ORGANIZATION_BLOCK "PullOrPlugOfModules"   // OB83, LAD, PullOrPlugOfModules
{ S7_Optimized_Access := 'TRUE' }
VERSION : 0.1
// stored: IsIECCheckEnabled false, SetENOAutomatically false
   VAR_INPUT
      LADDR : HW_IO;   // Hardware identifier
      Event_Class : Byte;   // 16#38/39: module inserted, removed
      Fault_ID : Byte;   // Fault identifier
   END_VAR
BEGIN
END_ORGANIZATION_BLOCK

ORGANIZATION_BLOCK "RackOrStationFailure"   // OB86, LAD, RackOrStationFailure
{ S7_Optimized_Access := 'TRUE' }
VERSION : 0.1
// stored: IsIECCheckEnabled false, SetENOAutomatically false
   VAR_INPUT
      LADDR : HW_DEVICE;   // Hardware identifier
      Event_Class : Byte;   // Event class
      Fault_ID : Byte;   // Fault identifier
   END_VAR
BEGIN
END_ORGANIZATION_BLOCK

FUNCTION "ByteArrayToString" : String   // FC15, SCL
{ S7_Optimized_Access := 'TRUE' }
VERSION : 0.1
// stored: AutoNumber true, IsIECCheckEnabled false, SetENOAutomatically false, UDAEnableTagReadback false
   VAR_INPUT
      Lenght : Int;
      ByteArray : Array[0..1024] of Byte;
   END_VAR
   VAR_OUTPUT
      ByteArrayToString_1 : String;
      ByteArrayToString_2 : String;
      ByteArrayToString_3 : String;
      ByteArrayToString_4 : String;
      ByteArrayToString_5 : String;
   END_VAR
   VAR_TEMP
      tempStr_1 : String;
      tempStr_2 : String;
      tempStr_3 : String;
      tempStr_4 : String;
      tempStr_5 : String;
      tempStr_6 : String;
      foundPos : Int;
      i : Int;
   END_VAR
BEGIN
   //STRING 1
   #tempStr_1 := '';
   FOR #i := 0 TO MIN(IN1 := #Lenght - 1, IN2 := 254) DO
       IF #ByteArray[#i] <> 0 THEN
           #tempStr_1 := CONCAT(IN1 := #tempStr_1, IN2 := CHAR_TO_STRING(BYTE_TO_CHAR(#ByteArray[#i])));
       END_IF;
   END_FOR;

   //STRING 2
   #tempStr_2 := '';
   FOR #i := 100 TO MIN(IN1 := #Lenght - 1, IN2 := 354) DO
       IF #ByteArray[#i] <> 0 THEN
           #tempStr_2 := CONCAT(IN1 := #tempStr_2, IN2 := CHAR_TO_STRING(BYTE_TO_CHAR(#ByteArray[#i])));
       END_IF;
   END_FOR;

   //STRING 3
   #tempStr_3 := '';
   FOR #i := 200 TO MIN(IN1 := #Lenght - 1, IN2 := 454) DO
       IF #ByteArray[#i] <> 0 THEN
           #tempStr_3 := CONCAT(IN1 := #tempStr_3, IN2 := CHAR_TO_STRING(BYTE_TO_CHAR(#ByteArray[#i])));
       END_IF;
   END_FOR;

   //STRING 4
   #tempStr_4 := '';
   FOR #i := 300 TO MIN(IN1 := #Lenght - 1, IN2 := 554) DO
       IF #ByteArray[#i] <> 0 THEN
           #tempStr_4 := CONCAT(IN1 := #tempStr_4, IN2 := CHAR_TO_STRING(BYTE_TO_CHAR(#ByteArray[#i])));
       END_IF;
   END_FOR;

   // //STRING 5
   #tempStr_5 := '';
   FOR #i := 400 TO MIN(IN1 := #Lenght - 1, IN2 := 654) DO
       IF #ByteArray[#i] <> 0 THEN
           #tempStr_5 := CONCAT(IN1 := #tempStr_5, IN2 := CHAR_TO_STRING(BYTE_TO_CHAR(#ByteArray[#i])));
       END_IF;
   END_FOR;

   // //STRING 6
   #tempStr_6 := '';
   FOR #i := 500 TO MIN(IN1 := #Lenght - 1, IN2 := 763) DO
       IF #ByteArray[#i] <> 0 THEN
           #tempStr_6 := CONCAT(IN1 := #tempStr_6, IN2 := CHAR_TO_STRING(BYTE_TO_CHAR(#ByteArray[#i])));
       END_IF;
   END_FOR;

   // Remove '$R$L'
   // string 1
   #foundPos := FIND(IN1 := #tempStr_1, IN2 := '$R$L');
   WHILE #foundPos > 0 DO
       #tempStr_1 := REPLACE(IN1 := #tempStr_1, IN2 := '', P := #foundPos, L := 2);
       #foundPos := FIND(IN1 := #tempStr_1, IN2 := '$R$L');
   END_WHILE;

   // string 2
   #foundPos := FIND(IN1 := #tempStr_2, IN2 := '$R$L');
   WHILE #foundPos > 0 DO
       #tempStr_2 := REPLACE(IN1 := #tempStr_2, IN2 := '', P := #foundPos, L := 2);
       #foundPos := FIND(IN1 := #tempStr_2, IN2 := '$R$L');
   END_WHILE;

   // string 3
   #foundPos := FIND(IN1 := #tempStr_3, IN2 := '$R$L');
   WHILE #foundPos > 0 DO
       #tempStr_3 := REPLACE(IN1 := #tempStr_3, IN2 := '', P := #foundPos, L := 2);
       #foundPos := FIND(IN1 := #tempStr_3, IN2 := '$R$L');
   END_WHILE;

   // string 4
   #foundPos := FIND(IN1 := #tempStr_4, IN2 := '$R$L');
   WHILE #foundPos > 0 DO
       #tempStr_4 := REPLACE(IN1 := #tempStr_4, IN2 := '', P := #foundPos, L := 2);
       #foundPos := FIND(IN1 := #tempStr_4, IN2 := '$R$L');
   END_WHILE;

   // string 5
   #foundPos := FIND(IN1 := #tempStr_5, IN2 := '$R$L');
   WHILE #foundPos > 0 DO
       #tempStr_5 := REPLACE(IN1 := #tempStr_5, IN2 := '', P := #foundPos, L := 2);
       #foundPos := FIND(IN1 := #tempStr_5, IN2 := '$R$L');
   END_WHILE;

   // string 6
   #foundPos := FIND(IN1 := #tempStr_6, IN2 := '$R$L');
   WHILE #foundPos > 0 DO
       #tempStr_6 := REPLACE(IN1 := #tempStr_6, IN2 := '', P := #foundPos, L := 2);
       #foundPos := FIND(IN1 := #tempStr_6, IN2 := '$R$L');
   END_WHILE;

   #ByteArrayToString := #tempStr_1;
   #ByteArrayToString_1 := #tempStr_2;
   #ByteArrayToString_2 := #tempStr_3;
   #ByteArrayToString_3 := #tempStr_4;
   #ByteArrayToString_4 := #tempStr_5;
   #ByteArrayToString_5 := #tempStr_6;
END_FUNCTION

FUNCTION "ByteArrayToString_1" : String   // FC23, SCL
{ S7_Optimized_Access := 'TRUE' }
VERSION : 0.1
// stored: AutoNumber true, IsIECCheckEnabled false, SetENOAutomatically false, UDAEnableTagReadback false
   VAR_INPUT
      Lenght : Int;
      ByteArray : Array[1..200] of Byte;
   END_VAR
   VAR_TEMP
      tempStr_1 : String;
      foundPos : Int;
      i : Int;
   END_VAR
BEGIN
   #tempStr_1 := '';
   FOR #i := 1 TO MIN(IN1 := #Lenght - 1, IN2 := 200) DO
       IF #ByteArray[#i] <> 0 THEN
           #tempStr_1 := CONCAT(IN1 := #tempStr_1, IN2 := CHAR_TO_STRING(BYTE_TO_CHAR(#ByteArray[#i])));
       END_IF;
   END_FOR;

   // Remove '$02'
   // string 1
   #foundPos := FIND(IN1 := #tempStr_1, IN2 := '$02');
   WHILE #foundPos > 0 DO
       #tempStr_1 := REPLACE(IN1 := #tempStr_1, IN2 := '', P := #foundPos, L := 1);
       #foundPos := FIND(IN1 := #tempStr_1, IN2 := '$02');
   END_WHILE;

   #ByteArrayToString_1 := #tempStr_1;
END_FUNCTION

FUNCTION "CharsArrayToString" : String   // FC27, SCL
{ S7_Optimized_Access := 'TRUE' }
VERSION : 0.1
// stored: AutoNumber true, IsIECCheckEnabled false, SetENOAutomatically false, UDAEnableTagReadback false
   VAR_INPUT
      Lenght : Int;
      CharsArray : Array[1..16] of Char;
   END_VAR
   VAR_TEMP
      tempStr_1 : String;
      foundPos : Int;
      i : Int;
   END_VAR
BEGIN
   #tempStr_1 := '';
   FOR #i := 1 TO MIN(IN1 := #Lenght - 1, IN2 := 16) DO
       IF #CharsArray[#i] <> '$00' THEN
           #tempStr_1 := CONCAT(IN1 := #tempStr_1, IN2 := CHAR_TO_STRING(#CharsArray[#i]));
       END_IF;
   END_FOR;

   // Remove '$00'
   // string 1
   #foundPos := FIND(IN1 := #tempStr_1, IN2 := '$00');
   WHILE #foundPos > 0 DO
       #tempStr_1 := REPLACE(IN1 := #tempStr_1, IN2 := '', P := #foundPos, L := 1);
       #foundPos := FIND(IN1 := #tempStr_1, IN2 := '$00');
   END_WHILE;

   #CharsArrayToString := #tempStr_1;
END_FUNCTION

FUNCTION "FindBoolField" : Bool   // FC17, SCL
{ S7_Optimized_Access := 'TRUE' }
VERSION : 0.1
// stored: AutoNumber true, IsIECCheckEnabled false, SetENOAutomatically false, UDAEnableTagReadback false
   VAR_INPUT
      FieldName : String;
      JsonStr : String;
   END_VAR
   VAR_TEMP
      searchStr : String;
      foundPos : Int;
      valueStr : String;
      afterField : String;
      bResult : Bool;
   END_VAR
BEGIN
   // Build search string
   #searchStr := CONCAT(IN1 := '"', IN2 := #FieldName);
   #searchStr := CONCAT(IN1 := #searchStr, IN2 := '" :');

   // Serach for JSON field
   #foundPos := FIND(IN1 := #JsonStr, IN2 := #searchStr);

   IF #foundPos > 0 THEN
       // Take to 20 characters after the field
       #afterField := MID(IN := #JsonStr, P := #foundPos + LEN(#searchStr), L := 20);

       // Normalize to remove whitespace if necessary
       // (or compare directly)
       IF FIND(IN1 := #afterField, IN2 := 'true') > 0 THEN
           #bResult := TRUE;
       ELSIF FIND(IN1 := #afterField, IN2 := 'false') > 0 THEN
           #bResult := FALSE;
       ELSE
           #bResult := FALSE; // default if value not found
       END_IF;
   ELSE
       #bResult := FALSE;
   END_IF;

   #FindBoolField := #bResult;
END_FUNCTION

FUNCTION "FindDINTFieldFragmented" : DInt   // FC20, SCL
{ S7_Optimized_Access := 'TRUE' }
VERSION : 0.1
// stored: AutoNumber true, IsIECCheckEnabled false, SetENOAutomatically false, UDAEnableTagReadback false
   VAR_INPUT
      FieldName : String;
      Str1 : String;
      Str2 : String;
   END_VAR
   VAR_TEMP
      searchStr : String;
      iStart : Int;
      iEnd : Int;
      tempVal : String;
      fieldFound : Bool;
      loopIdx : Int;
   END_VAR
BEGIN
   // Build search string
   #searchStr := CONCAT(IN1 := '"', IN2 := #FieldName);
   #searchStr := CONCAT(IN1 := #searchStr, IN2 := '" :');

   // Serach for JSON field
   #iStart := FIND(IN1 := #Str1, IN2 := #searchStr);

   IF #iStart > 0 THEN
       // Found full field in String_1
       #iEnd := FIND(IN1 := MID(IN := #Str1, P := #iStart + LEN(#searchStr), L := 20), IN2 := ',');
       IF #iEnd = 0 THEN
           #iEnd := FIND(IN1 := MID(IN := #Str1, P := #iStart + LEN(#searchStr), L := 20), IN2 := '}');
       END_IF;
       IF #iEnd > 0 THEN
           #tempVal := MID(IN := #Str1, P := #iStart + LEN(#searchStr), L := #iEnd - 1);
           #fieldFound := TRUE;
       END_IF;
   END_IF;

   // Search for full field in Str2
   IF NOT #fieldFound THEN
       #iStart := FIND(IN1 := #Str2, IN2 := #searchStr);
       IF #iStart > 0 THEN
           #iEnd := FIND(IN1 := MID(IN := #Str2, P := #iStart + LEN(#searchStr), L := 20), IN2 := ',');
           IF #iEnd = 0 THEN
               #iEnd := FIND(IN1 := MID(IN := #Str2, P := #iStart + LEN(#searchStr), L := 20), IN2 := '}');
           END_IF;
           IF #iEnd > 0 THEN
               #tempVal := MID(IN := #Str2, P := #iStart + LEN(#searchStr), L := #iEnd - 1);
               #fieldFound := TRUE;
           END_IF;
       END_IF;
   END_IF;

   // Search for fragmented field: end of name in Str1 and beginning in Str2
   IF NOT #fieldFound THEN
       // Examines last 10 characters of String_1
       FOR #loopIdx := LEN(#Str1) - 15 TO LEN(#Str1) DO
           IF MID(IN := #Str1, P := #loopIdx, L := 1) = '"' THEN
               #tempVal := MID(IN := #Str1, P := #loopIdx, L := LEN(#Str1) - #loopIdx + 1);
               #tempVal := CONCAT(IN1 := #tempVal, IN2 := #Str2); // concatenates piece from beginning of String_2
               #iStart := FIND(IN1 := #tempVal, IN2 := #searchStr);
               IF #iStart > 0 THEN
                   #iEnd := FIND(IN1 := MID(IN := #tempVal, P := #iStart + LEN(#searchStr), L := 20), IN2 := ',');
                   IF #iEnd = 0 THEN
                       #iEnd := FIND(IN1 := MID(IN := #tempVal, P := #iStart + LEN(#searchStr), L := 20), IN2 := '}');
                   END_IF;
                   IF #iEnd > 0 THEN
                       #tempVal := MID(IN := #tempVal, P := #iStart + LEN(#searchStr), L := #iEnd - 1);
                       #fieldFound := TRUE;
                   END_IF;
               END_IF;
               EXIT; // found, you can leave
           END_IF;
       END_FOR;
   END_IF;

   // Return value
   IF #fieldFound THEN
       #FindDINTFieldFragmented := STRING_TO_DINT(#tempVal);
   ELSE
       #FindDINTFieldFragmented := -9999; // default value if not found
   END_IF;
END_FUNCTION

FUNCTION "FindINTFieldFragmented" : Int   // FC22, SCL
{ S7_Optimized_Access := 'TRUE' }
VERSION : 0.1
// stored: AutoNumber true, IsIECCheckEnabled false, SetENOAutomatically false, UDAEnableTagReadback false
   VAR_INPUT
      FieldName : String;
      Str1 : String;
      Str2 : String;
   END_VAR
   VAR_TEMP
      searchStr : String;
      iStart : Int;
      iEnd : Int;
      tempVal : String;
      fieldFound : Bool;
      loopIdx : Int;
   END_VAR
BEGIN
   // Build search string
   #searchStr := CONCAT(IN1 := '"', IN2 := #FieldName);
   #searchStr := CONCAT(IN1 := #searchStr, IN2 := '" :');

   // Serach for JSON field
   #iStart := FIND(IN1 := #Str1, IN2 := #searchStr);

   IF #iStart > 0 THEN
       // Found full field in String_1
       #iEnd := FIND(IN1 := MID(IN := #Str1, P := #iStart + LEN(#searchStr), L := 20), IN2 := ',');
       IF #iEnd = 0 THEN
           #iEnd := FIND(IN1 := MID(IN := #Str1, P := #iStart + LEN(#searchStr), L := 20), IN2 := '}');
       END_IF;
       IF #iEnd > 0 THEN
           #tempVal := MID(IN := #Str1, P := #iStart + LEN(#searchStr), L := #iEnd - 1);
           #fieldFound := TRUE;
       END_IF;
   END_IF;

   // Search for full field in Str2
   IF NOT #fieldFound THEN
       #iStart := FIND(IN1 := #Str2, IN2 := #searchStr);
       IF #iStart > 0 THEN
           #iEnd := FIND(IN1 := MID(IN := #Str2, P := #iStart + LEN(#searchStr), L := 20), IN2 := ',');
           IF #iEnd = 0 THEN
               #iEnd := FIND(IN1 := MID(IN := #Str2, P := #iStart + LEN(#searchStr), L := 20), IN2 := '}');
           END_IF;
           IF #iEnd > 0 THEN
               #tempVal := MID(IN := #Str2, P := #iStart + LEN(#searchStr), L := #iEnd - 1);
               #fieldFound := TRUE;
           END_IF;
       END_IF;
   END_IF;

   // Search for fragmented field: end of name in Str1 and beginning in Str2
   IF NOT #fieldFound THEN
       // Examines last 10 characters of String_1
       FOR #loopIdx := LEN(#Str1) - 15 TO LEN(#Str1) DO
           IF MID(IN := #Str1, P := #loopIdx, L := 1) = '"' THEN
               #tempVal := MID(IN := #Str1, P := #loopIdx, L := LEN(#Str1) - #loopIdx + 1);
               #tempVal := CONCAT(IN1 := #tempVal, IN2 := #Str2); // concatenates piece from beginning of String_2
               #iStart := FIND(IN1 := #tempVal, IN2 := #searchStr);
               IF #iStart > 0 THEN
                   #iEnd := FIND(IN1 := MID(IN := #tempVal, P := #iStart + LEN(#searchStr), L := 20), IN2 := ',');
                   IF #iEnd = 0 THEN
                       #iEnd := FIND(IN1 := MID(IN := #tempVal, P := #iStart + LEN(#searchStr), L := 20), IN2 := '}');
                   END_IF;
                   IF #iEnd > 0 THEN
                       #tempVal := MID(IN := #tempVal, P := #iStart + LEN(#searchStr), L := #iEnd - 1);
                       #fieldFound := TRUE;
                   END_IF;
               END_IF;
               EXIT; // found, you can leave
           END_IF;
       END_FOR;
   END_IF;

   // Return value
   IF #fieldFound THEN
       #FindINTFieldFragmented := STRING_TO_INT(#tempVal);
   ELSE
       #FindINTFieldFragmented := -9999; // default value if not found
   END_IF;
END_FUNCTION

FUNCTION "FindIntField" : Int   // FC18, SCL
{ S7_Optimized_Access := 'TRUE' }
VERSION : 0.1
// stored: AutoNumber true, IsIECCheckEnabled false, SetENOAutomatically false, UDAEnableTagReadback false
   VAR_INPUT
      FieldName : String;
      JsonStr : String;
   END_VAR
   VAR_TEMP
      searchStr : String;
      foundPos : Int;
      valueStr : String;
      delimPos : Int;
   END_VAR
BEGIN
   // Set up the search pattern, e.g. '"id":'
   #searchStr := CONCAT(IN1 := '"', IN2 := #FieldName);
   #searchStr := CONCAT(IN1 := #searchStr, IN2 := '" :');

   // Search the field
   #foundPos := FIND(IN1 := #JsonStr, IN2 := #searchStr);

   IF #foundPos > 0 THEN
       // Try to find a comma after the value
       #delimPos := FIND(
                         IN1 := MID(IN := #JsonStr, P := #foundPos + LEN(#searchStr), L := 10),
                         IN2 := ','
       );

       // If there is no comma, try to find the closing brace '}'
       IF #delimPos = 0 THEN
           #delimPos := FIND(
                             IN1 := MID(IN := #JsonStr, P := #foundPos + LEN(#searchStr), L := 10),
                             IN2 := '}'
           );
       END_IF;

       // If you find the end of value, extract the value
       IF #delimPos > 0 THEN
           #valueStr := MID(
                            IN := #JsonStr,
                            P := #foundPos + LEN(#searchStr),
                            L := #delimPos - 1
           );
           #FindIntField := STRING_TO_INT(#valueStr);
           RETURN;
       END_IF;
   END_IF;

   // Default return if not found or error
   #FindIntField := -9999;
END_FUNCTION

FUNCTION "FindSTRINGFieldFragmented" : String   // FC21, SCL
{ S7_Optimized_Access := 'TRUE' }
VERSION : 0.1
// stored: AutoNumber true, IsIECCheckEnabled false, SetENOAutomatically false, UDAEnableTagReadback false
   VAR_INPUT
      FieldName : String;
      Str1 : String;
      Str2 : String;
   END_VAR
   VAR_TEMP
      searchStr : String;
      iStart : Int;
      iEnd : Int;
      tempVal : String;
      fieldFound : Bool;
      loopIdx : Int;
   END_VAR
BEGIN
   // Build search string
   #searchStr := CONCAT(IN1 := '"', IN2 := #FieldName);
   #searchStr := CONCAT(IN1 := #searchStr, IN2 := '" :');

   // Serach for JSON field
   #iStart := FIND(IN1 := #Str1, IN2 := #searchStr);

   IF #iStart > 0 THEN
       // Found full field in String_1
       #iEnd := FIND(IN1 := MID(IN := #Str1, P := #iStart + LEN(#searchStr), L := 20), IN2 := ',');
       IF #iEnd = 0 THEN
           #iEnd := FIND(IN1 := MID(IN := #Str1, P := #iStart + LEN(#searchStr), L := 20), IN2 := '}');
       END_IF;
       IF #iEnd > 0 THEN
           #tempVal := MID(IN := #Str1, P := #iStart + LEN(#searchStr), L := #iEnd - 1);
           #fieldFound := TRUE;
       END_IF;
   END_IF;

   // Search for full field in Str2
   IF NOT #fieldFound THEN
       #iStart := FIND(IN1 := #Str2, IN2 := #searchStr);
       IF #iStart > 0 THEN
           #iEnd := FIND(IN1 := MID(IN := #Str2, P := #iStart + LEN(#searchStr), L := 20), IN2 := ',');
           IF #iEnd = 0 THEN
               #iEnd := FIND(IN1 := MID(IN := #Str2, P := #iStart + LEN(#searchStr), L := 20), IN2 := '}');
           END_IF;
           IF #iEnd > 0 THEN
               #tempVal := MID(IN := #Str2, P := #iStart + LEN(#searchStr), L := #iEnd - 1);
               #fieldFound := TRUE;
           END_IF;
       END_IF;
   END_IF;

   // Search for fragmented field: end of name in Str1 and beginning in Str2
   IF NOT #fieldFound THEN
       // Examines last 10 characters of String_1
       FOR #loopIdx := LEN(#Str1) - 15 TO LEN(#Str1) DO
           IF MID(IN := #Str1, P := #loopIdx, L := 1) = '"' THEN
               #tempVal := MID(IN := #Str1, P := #loopIdx, L := LEN(#Str1) - #loopIdx + 1);
               #tempVal := CONCAT(IN1 := #tempVal, IN2 := #Str2); // concatenates piece from beginning of String_2
               #iStart := FIND(IN1 := #tempVal, IN2 := #searchStr);
               IF #iStart > 0 THEN
                   #iEnd := FIND(IN1 := MID(IN := #tempVal, P := #iStart + LEN(#searchStr), L := 20), IN2 := ',');
                   IF #iEnd = 0 THEN
                       #iEnd := FIND(IN1 := MID(IN := #tempVal, P := #iStart + LEN(#searchStr), L := 20), IN2 := '}');
                   END_IF;
                   IF #iEnd > 0 THEN
                       #tempVal := MID(IN := #tempVal, P := #iStart + LEN(#searchStr), L := #iEnd - 1);
                       #fieldFound := TRUE;
                   END_IF;
               END_IF;
               EXIT; // found, you can leave
           END_IF;
       END_FOR;
   END_IF;

   // Return value
   IF #fieldFound THEN
       #FindSTRINGFieldFragmented := #tempVal;
   ELSE
       #FindSTRINGFieldFragmented := 'NOT FOUND'; // default value if not found
   END_IF;
END_FUNCTION

FUNCTION "FindStringField" : String   // FC19, SCL
{ S7_Optimized_Access := 'TRUE' }
VERSION : 0.1
// stored: AutoNumber true, IsIECCheckEnabled false, SetENOAutomatically false, UDAEnableTagReadback false
   VAR_INPUT
      FieldName : String;
      JsonStr : String;
   END_VAR
   VAR_TEMP
      searchStr : String;
      foundPos : Int;
      resultStr : String;
      quotePos1 : Int;
      quotePos2 : Int;
   END_VAR
BEGIN
   // Sets search pattern → ex: '"loadstate":'
   #searchStr := CONCAT(IN1 := '"', IN2 := #FieldName);
   #searchStr := CONCAT(IN1 := #searchStr, IN2 := '" :');

   // Search in JSON
   #foundPos := FIND(IN1 := #JsonStr, IN2 := #searchStr);

   IF #foundPos > 0 THEN
       // Finds first quote after field
       #quotePos1 := FIND(IN1 := MID(IN := #JsonStr, P := #foundPos + LEN(#searchStr), L := 20), IN2 := '"');

       IF #quotePos1 > 0 THEN
           // Finds second quote after the first
           #quotePos2 := FIND(
                              IN1 := MID(IN := #JsonStr, P := #foundPos + LEN(IN := #searchStr) + #quotePos1, L := 10),
                              IN2 := '"'
           );

           IF #quotePos2 > 0 THEN
               #resultStr := MID(
                                 IN := #JsonStr,
                                 P := #foundPos + LEN(#searchStr) + #quotePos1,
                                 L := #quotePos2 - 1
               );
               #FindStringField := #resultStr;
               RETURN;
           END_IF;
       END_IF;
   END_IF;

   // If not found, returns empty string
   #FindStringField := '';
END_FUNCTION

FUNCTION "ID_Decode_F" : Void   // FC3, SCL
{ S7_Optimized_Access := 'TRUE' }
VERSION : 0.1
// stored: AutoNumber true, IsIECCheckEnabled false, SetENOAutomatically false, UDAEnableTagReadback false
   VAR_INPUT
      ID : DInt;
   END_VAR
   VAR_IN_OUT
      ID_Decoded : "ID_Decoded";
   END_VAR
   VAR_TEMP
      Temp : UInt;
   END_VAR
BEGIN

   // Extract XX (first two digits)
   #ID_Decoded.Device_Type := #ID / 10000;        // 123456 / 10000 = 12

   // Extract YY (middle two digits)
   #ID_Decoded.Level := (#ID MOD 10000) / 100; // 123456 % 10000 = 3456 → 3456 / 100 = 34

   // Extract ZZ (last two digits)
   #ID_Decoded.VTD := #ID MOD 100;       // 123456 % 100 = 56
END_FUNCTION

FUNCTION "IsIPAddress" : Bool   // FC4, SCL
TITLE = IsIPAddress
{ S7_Optimized_Access := 'TRUE' }
VERSION : 0.1
// Evaluates whether a given String contains a valid IP address
// stored: AutoNumber true, IsIECCheckEnabled true, SetENOAutomatically true, UDAEnableTagReadback false
   VAR_INPUT
      address : String;   // Address to be evaluated
   END_VAR
   VAR_OUTPUT
      ipAddress : IP_V4;   // Parsed IP address if passed address is IP address
   END_VAR
   VAR_TEMP
      tempAddress : String;   // Passed address
      tempOctet : String;   // Current octet
      tempIndex : DInt;   // Index for loop
      tempPos : Int;   // Position of found separator
      tempNum : Int;   // Converted octet
      tempIp : IP_V4;   // Parsed IP address
   END_VAR
   VAR CONSTANT
      MAX_VALUE : USInt := 255;   // Max. valid value of octet
      NUM_OCTETS : DInt := 4;   // Number of octets
      CHAR_ZERO : Char := '0';   // ASCII character '0'
   END_VAR
   // Ret_Val : Return value
BEGIN
   REGION BLOCK INFO HEADER
     //===============================================================================
     // SIEMENS / (c)Copyright 2024
     //-------------------------------------------------------------------------------
     // Title:        IsIPAddress
     // Function:     Evaluates whether a given String contains a valid IP address
     // Library:      --
     // Author:       Siemens Industry Online Support
     // Tested with:  CPU 1515-2 PN V3.1
     // Engineering:  TIA Portal V17
     // Restrictions: --
     // Requirements: S7-1200 with firmware V4.4 or higher
     //               S7-1500 with firmware V2.0 or higher
     //-------------------------------------------------------------------------------
     // Change log table:
     // Version  | Date       | Expert in charge       | Changes applied
     //-------------------------------------------------------------------------------
     // 01.00.00 | 2024-02-12 | Online Support         | First released version
     //===============================================================================
   END_REGION

   #tempAddress := #address;
   #IsIPAddress := FALSE; // Will be overwritten if IP address is detected
   #ipAddress := #tempIp; // Zero output parameter

   FOR #tempIndex := 1 TO #NUM_OCTETS DO
     #tempPos := FIND(IN1 := #tempAddress, IN2 := '.'); // Find separator

     IF (#tempPos > 0 OR #tempIndex = #NUM_OCTETS) // Separator found with exception of last octet
       AND NOT (#tempPos > 0 AND #tempIndex = #NUM_OCTETS) // No separator found in last octet
       AND #tempPos <= 4 // 3  characters or less
     THEN
       IF #tempIndex < #NUM_OCTETS THEN // First three octets
         #tempOctet := LEFT(IN := #tempAddress, L := #tempPos - 1);
       ELSE// Last octet
         #tempOctet := #tempAddress;
       END_IF;

       STRG_VAL(IN := #tempOctet,
                FORMAT := 0,
                P := 1,
                OUT => #tempNum);

       IF #tempNum >= 0 AND #tempNum <= #MAX_VALUE // Within 0 and 255
         AND NOT (#tempNum = 0 AND #tempIndex = 1) // Not 0 in first octet
         AND NOT (#tempNum = 0 AND #tempOctet[1] <> #CHAR_ZERO) // Not 0 because of invalid character
       THEN
         #tempIp.ADDR[#tempIndex] := INT_TO_BYTE(#tempNum);
         #tempAddress := RIGHT(IN := #tempAddress, L := LEN(#tempAddress) - #tempPos); // Remove evaluated octet
       ELSE // Address is not IP address
         EXIT;
       END_IF;
     ELSE // Address is not IP address
       EXIT;
     END_IF;

     IF #tempIndex = #NUM_OCTETS THEN // End of loop reached, address is IP address
       #ipAddress := #tempIp;
       #IsIPAddress := true;
     END_IF;
   END_FOR;
END_FUNCTION

FUNCTION "LMQTT_ConvertToUtf8" : Void   // FC6, SCL
TITLE = LMQTT_ConvertToUtf8
{ S7_Optimized_Access := 'TRUE' }
AUTHOR : SIEMENS
FAMILY : LMQTT
VERSION : 1.0
// Function to convert a WCHAR to a UTF-8 conformant byte sequence
// stored: AutoNumber true, IsIECCheckEnabled true, SetENOAutomatically false, UDAEnableTagReadback false
   VAR_INPUT
      character : WChar;   // Character that shall be converted to UTF-8
   END_VAR
   VAR_OUTPUT
      convertedUtf8 : DWord;   // UTF-8 conformant byte sequence. B0 stores first Byte, B1 second and B2 third Byte. B3 is not used
      bytesUsed : USInt;   // Amount of Bytes converted. Ranges from 1 to 3.
      error : Bool;   // TRUE: An error occurred during the execution of the FC
      status : Word;   // 16#0000 - 16#7FFF: Status of the FC, 16#8000 - 16#FFFF: Error identification
   END_VAR
   VAR_TEMP
      tempStatus : Word;   // temp value for output 'status'
      tempConvertedUtf8 : DWord;   // temp value for output 'convertedUtf8'
      tempBytesUsed : USInt;   // temp value for output 'bytesUsed'
      tempCharacter : WChar;   // temp value for input 'character'
   END_VAR
   VAR CONSTANT
      STATUS_NO_ERROR : Word := 16#0000;   // no error status
      STATUS_EXECUTION_FINISHED : Word := 16#0000;   // Execution finished without errors
      ERR_UNDEFINED : Word := 16#8000;   // Error due to an undefined case
      USINT_NULL : USInt := 0;   // Init value with 0
      DWORD_NULL : DWord := 16#0000_0000;   // Init value with 0
      EMPTY_WCHAR : WChar := WCHAR#' ';   // Empty WChar for comparison
      BELOW_7F : Word := 16#007F;   // Upper limit for character if only one Byte used
      BELOW_7FF : Word := 16#07FF;   // Upper limit for character if two Byte used
      BELOW_MAX_FFFF : Word := 16#FFFF;   // Upper limit for character if three Byte used
      BYTE_3F : Byte := 16#3F;   // Conversion Value
      BYTE_80 : Byte := 16#80;   // Conversion Value
      BYTE_C0 : Byte := 16#C0;   // Conversion Value
      BYTE_E0 : Byte := 16#E0;   // Conversion Value
      USINT_ONE : USInt := 1;   // Const Value to assign amount of bytes used
      USINT_TWO : USInt := 2;   // Const Value to assign amount of bytes used
      USINT_THREE : USInt := 3;   // Const Value to assign amount of bytes used
   END_VAR
   // Ret_Val : No return for this FC - see error and status output
BEGIN
   REGION BLOCK INFO HEADER
       //=============================================================================
       // SIEMENS AG
       // (c)Copyright 2020
       //-----------------------------------------------------------------------------
       // Library:       LMQTT
       // Tested with:   CPU 1516-3 PN/DP V2.8
       // Engineering:   TIA Portal V16
       // Restrictions:  --
       // Requirements:  --
       // Functionality: Converts a single WChar Character to a valid UTF-8 encoded byte sequence and saves this to a DWord.
       //                The amount of bytes saved is stored in bytesUsed Output.
       //-----------------------------------------------------------------------------
       // Change log table:
       // Version    Date         Expert in charge         Changes applied
       // 03.00.00   01.10.2020   Siemens Online Support   First released version
       //=============================================================================
   END_REGION

   REGION INITIALISATION  
       // Initialize functionality: reset of variables, diagnostics, etc.
       #tempConvertedUtf8 := #DWORD_NULL;
       #tempBytesUsed := #USINT_NULL;
       #tempStatus := #STATUS_NO_ERROR;
       //assign temp value from input:
        #tempCharacter := #character;

   END_REGION

   REGION PROGRAM LOGIC
       // Use this region for application specific code
       IF #tempCharacter = #EMPTY_WCHAR THEN
           //will be only 1 byte occupied
           #tempConvertedUtf8 := WCHAR_TO_DWORD(#tempCharacter);
           #tempBytesUsed := #USINT_ONE;
       ELSIF (WCHAR_TO_WORD(#tempCharacter) <= (#BELOW_7F)) THEN
           //will be only 1 byte occupied
           #tempConvertedUtf8 := WCHAR_TO_DWORD(#tempCharacter);
           #tempBytesUsed := #USINT_ONE;
       ELSIF (WCHAR_TO_WORD(#tempCharacter) <= (#BELOW_7FF)) THEN
           //will be 2 byte occupied
           #tempConvertedUtf8.%B1 := (WCHAR_TO_BYTE(#tempCharacter) AND #BYTE_3F) OR #BYTE_80;
           #tempConvertedUtf8.%B0 := WORD_TO_BYTE(SHR(IN := WCHAR_TO_WORD(#tempCharacter), N := 6)) OR #BYTE_C0;
           #tempBytesUsed := #USINT_TWO;
       ELSIF (WCHAR_TO_WORD(#tempCharacter) <= (#BELOW_MAX_FFFF)) THEN
           //will be 3 byte occupied
           #tempConvertedUtf8.%B2 := (WCHAR_TO_BYTE(#tempCharacter) AND #BYTE_3F) OR #BYTE_80;
           #tempConvertedUtf8.%B1 := (WORD_TO_BYTE(SHR(IN := WCHAR_TO_WORD(#tempCharacter), N := 6)) AND #BYTE_3F) OR #BYTE_80;
           #tempConvertedUtf8.%B0 := WORD_TO_BYTE(SHR(IN := WCHAR_TO_WORD(#tempCharacter), N := 12)) OR #BYTE_E0;
           #tempBytesUsed := #USINT_THREE;
       END_IF;
   END_REGION

   REGION OUTPUTS
       // Write application specific temp values to outputs
       #bytesUsed := #tempBytesUsed;
       #convertedUtf8 := #tempConvertedUtf8;
       // Write error and status
       #error := #tempStatus.%X15;
       #status := #tempStatus;
       // ENO mechanism is not used --> ENO := TRUE;
       ENO := TRUE;
   END_REGION
END_FUNCTION

FUNCTION_BLOCK "Main_Safety_RTG1"   // FB1, F_FBD
{ S7_Optimized_Access := 'TRUE' }
VERSION : 0.1
// stored: AutoNumber false, IsIECCheckEnabled false, UDAEnableTagReadback false
   VAR
      SAFETY_OK_VTD : Bool;
      SAFETY_OK_CAROUSEL : Bool;
      MAIN_PANEL_OK : Bool;
      REMOTE_PANEL_OK : Bool;
      "E-STOP_INBOUND_OK" : Bool;
      PICK_STATION_OK : Bool;
      data_Safe : DInt;
      "HMI_E-STOP" : Bool;
   END_VAR
BEGIN

REGION Network 1: SAFETY OK VTD
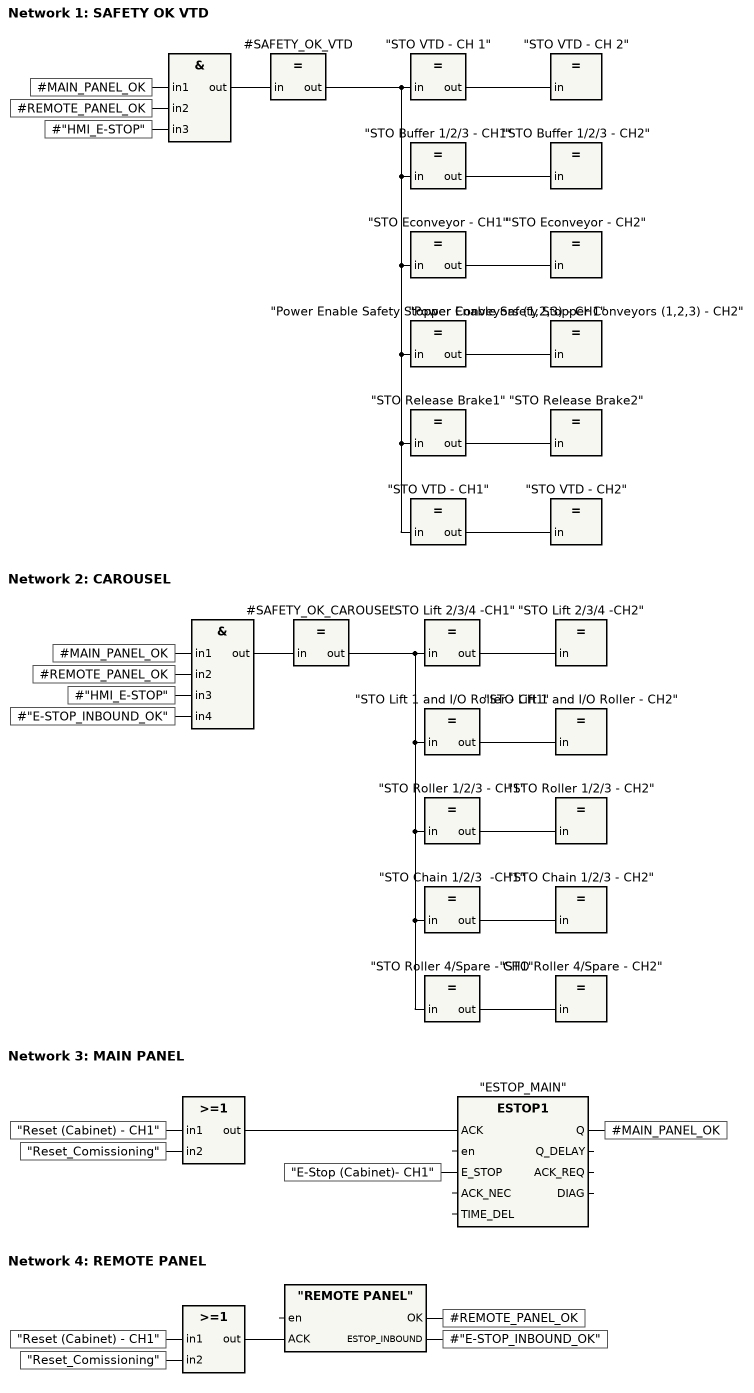
   #SAFETY_OK_VTD := #MAIN_PANEL_OK AND #REMOTE_PANEL_OK AND #"HMI_E-STOP";
   "STO VTD - CH 1" := #SAFETY_OK_VTD;
   "STO VTD - CH 2" := #SAFETY_OK_VTD;
   "STO Buffer 1/2/3 - CH1" := #SAFETY_OK_VTD;
   "STO Buffer 1/2/3 - CH2" := #SAFETY_OK_VTD;
   "STO Econveyor - CH1" := #SAFETY_OK_VTD;
   "STO Econveyor - CH2" := #SAFETY_OK_VTD;
   "Power Enable Safety Stopper Conveyors (1,2,3) - CH1" := #SAFETY_OK_VTD;
   "Power Enable Safety Stopper Conveyors (1,2,3) - CH2" := #SAFETY_OK_VTD;
   "STO Release Brake1" := #SAFETY_OK_VTD;
   "STO Release Brake2" := #SAFETY_OK_VTD;
   "STO VTD - CH1" := #SAFETY_OK_VTD;
   "STO VTD - CH2" := #SAFETY_OK_VTD;
END_REGION

REGION Network 2: CAROUSEL
   #SAFETY_OK_CAROUSEL := #MAIN_PANEL_OK AND #REMOTE_PANEL_OK AND #"HMI_E-STOP" AND #"E-STOP_INBOUND_OK";
   "STO Lift 2/3/4 -CH1" := #SAFETY_OK_CAROUSEL;
   "STO Lift 2/3/4 -CH2" := #SAFETY_OK_CAROUSEL;
   "STO Lift 1 and I/O Roller - CH1" := #SAFETY_OK_CAROUSEL;
   "STO Lift 1 and I/O Roller - CH2" := #SAFETY_OK_CAROUSEL;
   "STO Roller 1/2/3 - CH1" := #SAFETY_OK_CAROUSEL;
   "STO Roller 1/2/3 - CH2" := #SAFETY_OK_CAROUSEL;
   "STO Chain 1/2/3  -CH1" := #SAFETY_OK_CAROUSEL;
   "STO Chain 1/2/3 - CH2" := #SAFETY_OK_CAROUSEL;
   "STO Roller 4/Spare - CH1" := #SAFETY_OK_CAROUSEL;
   "STO Roller 4/Spare - CH2" := #SAFETY_OK_CAROUSEL;
END_REGION

REGION Network 3: MAIN PANEL
   "ESTOP_MAIN"(ACK := "Reset (Cabinet) - CH1" OR "Reset_Comissioning",   // ESTOP1
                E_STOP := "E-Stop (Cabinet)- CH1",
                Q => #MAIN_PANEL_OK);
END_REGION

REGION Network 4: REMOTE PANEL
   "REMOTE PANEL"(ACK := "Reset (Cabinet) - CH1" OR "Reset_Comissioning",
                  OK => #REMOTE_PANEL_OK,
                  ESTOP_INBOUND => #"E-STOP_INBOUND_OK");
END_REGION

REGION Network 5: 1=Acknowledgment for reintegration required
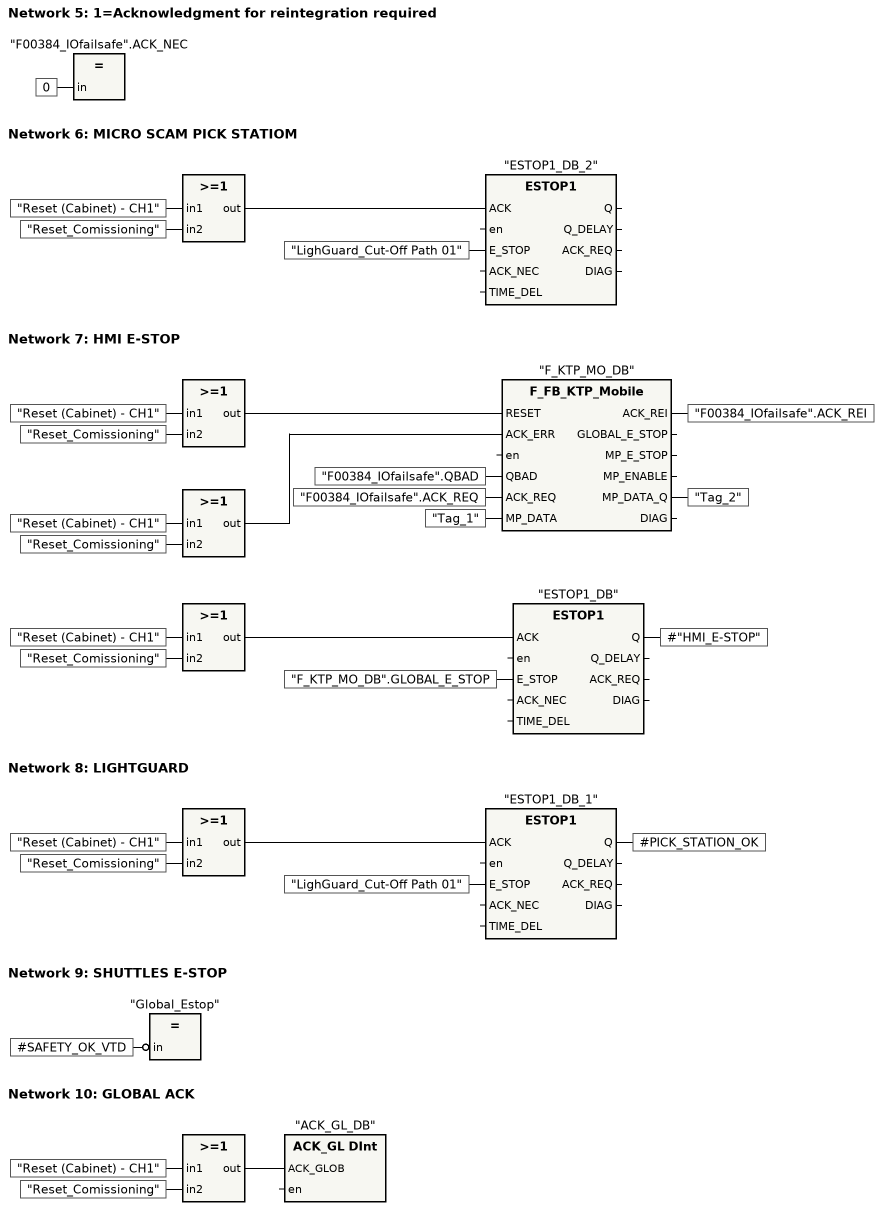
   "F00384_IOfailsafe".ACK_NEC := 0;
END_REGION

REGION Network 6: MICRO SCAM PICK STATIOM
   "ESTOP1_DB_2"(ACK := "Reset (Cabinet) - CH1" OR "Reset_Comissioning", E_STOP := "LighGuard_Cut-Off Path 01");   // ESTOP1
END_REGION

REGION Network 7: HMI E-STOP
   "F_KTP_MO_DB"(RESET := "Reset (Cabinet) - CH1" OR "Reset_Comissioning",   // F_FB_KTP_Mobile
                 ACK_ERR := "Reset (Cabinet) - CH1" OR "Reset_Comissioning",
                 QBAD := "F00384_IOfailsafe".QBAD,
                 ACK_REQ := "F00384_IOfailsafe".ACK_REQ,
                 MP_DATA := "Tag_1",
                 ACK_REI => "F00384_IOfailsafe".ACK_REI,
                 MP_DATA_Q => "Tag_2");
   "ESTOP1_DB"(ACK := "Reset (Cabinet) - CH1" OR "Reset_Comissioning",   // ESTOP1
               E_STOP := "F_KTP_MO_DB".GLOBAL_E_STOP,
               Q => #"HMI_E-STOP");
END_REGION

REGION Network 8: LIGHTGUARD
   "ESTOP1_DB_1"(ACK := "Reset (Cabinet) - CH1" OR "Reset_Comissioning",   // ESTOP1
                 E_STOP := "LighGuard_Cut-Off Path 01",
                 Q => #PICK_STATION_OK);
END_REGION

REGION Network 9: SHUTTLES E-STOP
   "Global_Estop" := NOT #SAFETY_OK_VTD;
END_REGION

REGION Network 10: GLOBAL ACK
   "ACK_GL_DB"(ACK_GLOB := "Reset (Cabinet) - CH1" OR "Reset_Comissioning");   // ACK_GL
END_REGION
END_FUNCTION_BLOCK

FUNCTION "REMOTE PANEL" : Void   // FC1, F_LAD
{ S7_Optimized_Access := 'TRUE' }
VERSION : 0.1
// stored: AutoNumber true, IsIECCheckEnabled false, UDAEnableTagReadback false
   VAR_INPUT
      ACK : Bool;
   END_VAR
   VAR_OUTPUT
      OK : Bool;
      ESTOP_INBOUND : Bool;
   END_VAR
BEGIN

REGION Network 1: REMOTE PANEL OK
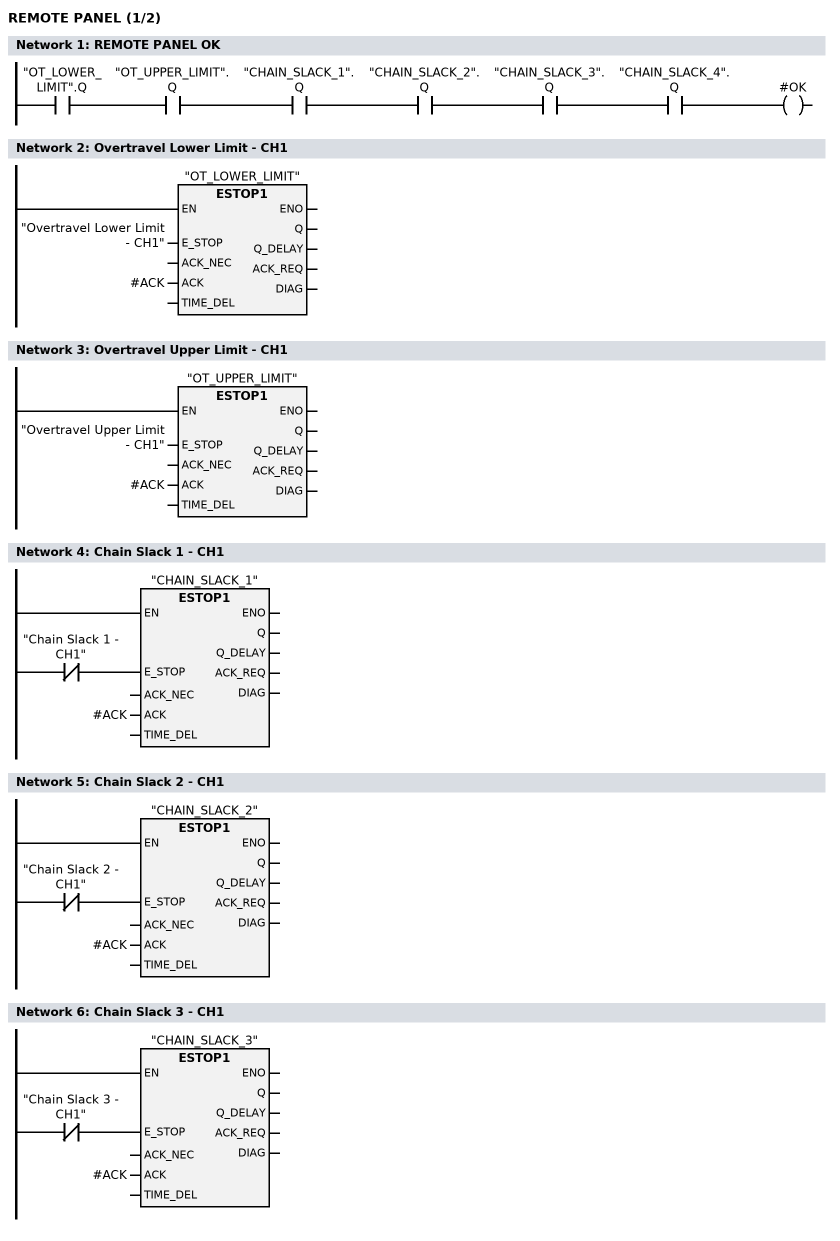
   RUNG wire#powerrail
      Contact( "OT_LOWER_LIMIT".Q )
      Contact( "OT_UPPER_LIMIT".Q )
      Contact( "CHAIN_SLACK_1".Q )
      Contact( "CHAIN_SLACK_2".Q )
      Contact( "CHAIN_SLACK_3".Q )
      Contact( "CHAIN_SLACK_4".Q )
      Coil( #OK )
   END_RUNG
   // the same network as SCL:
   #OK := "OT_LOWER_LIMIT".Q AND "OT_UPPER_LIMIT".Q AND "CHAIN_SLACK_1".Q AND "CHAIN_SLACK_2".Q AND "CHAIN_SLACK_3".Q AND "CHAIN_SLACK_4".Q;
END_REGION

REGION Network 2: Overtravel Lower Limit - CH1
   RUNG wire#powerrail
      "OT_LOWER_LIMIT".ESTOP1(E_STOP := "Overtravel Lower Limit - CH1", ACK_NEC :=, ACK := #ACK, TIME_DEL :=, Q =>, Q_DELAY =>, ACK_REQ =>, DIAG =>)
   END_RUNG
   // the same network as SCL:
   "OT_LOWER_LIMIT"(E_STOP := "Overtravel Lower Limit - CH1", ACK := #ACK);   // ESTOP1
END_REGION

REGION Network 3: Overtravel Upper Limit - CH1
   RUNG wire#powerrail
      "OT_UPPER_LIMIT".ESTOP1(E_STOP := "Overtravel Upper Limit - CH1", ACK_NEC :=, ACK := #ACK, TIME_DEL :=, Q =>, Q_DELAY =>, ACK_REQ =>, DIAG =>)
   END_RUNG
   // the same network as SCL:
   "OT_UPPER_LIMIT"(E_STOP := "Overtravel Upper Limit - CH1", ACK := #ACK);   // ESTOP1
END_REGION

REGION Network 4: Chain Slack 1 - CH1
   RUNG wire#powerrail
      "CHAIN_SLACK_1".ESTOP1(E_STOP := wire#w1, ACK_NEC :=, ACK := #ACK, TIME_DEL :=, Q =>, Q_DELAY =>, ACK_REQ =>, DIAG =>)
   END_RUNG
   RUNG wire#powerrail
      I_Contact( "Chain Slack 1 - CH1" )
   END_RUNG wire#w1
   // the same network as SCL:
   "CHAIN_SLACK_1"(E_STOP := NOT "Chain Slack 1 - CH1", ACK := #ACK);   // ESTOP1
END_REGION

REGION Network 5: Chain Slack 2 - CH1
   RUNG wire#powerrail
      "CHAIN_SLACK_2".ESTOP1(E_STOP := wire#w1, ACK_NEC :=, ACK := #ACK, TIME_DEL :=, Q =>, Q_DELAY =>, ACK_REQ =>, DIAG =>)
   END_RUNG
   RUNG wire#powerrail
      I_Contact( "Chain Slack 2 - CH1" )
   END_RUNG wire#w1
   // the same network as SCL:
   "CHAIN_SLACK_2"(E_STOP := NOT "Chain Slack 2 - CH1", ACK := #ACK);   // ESTOP1
END_REGION

REGION Network 6: Chain Slack 3 - CH1
   RUNG wire#powerrail
      "CHAIN_SLACK_3".ESTOP1(E_STOP := wire#w1, ACK_NEC :=, ACK := #ACK, TIME_DEL :=, Q =>, Q_DELAY =>, ACK_REQ =>, DIAG =>)
   END_RUNG
   RUNG wire#powerrail
      I_Contact( "Chain Slack 3 - CH1" )
   END_RUNG wire#w1
   // the same network as SCL:
   "CHAIN_SLACK_3"(E_STOP := NOT "Chain Slack 3 - CH1", ACK := #ACK);   // ESTOP1
END_REGION

REGION Network 7: Chain Slack 4 - CH1
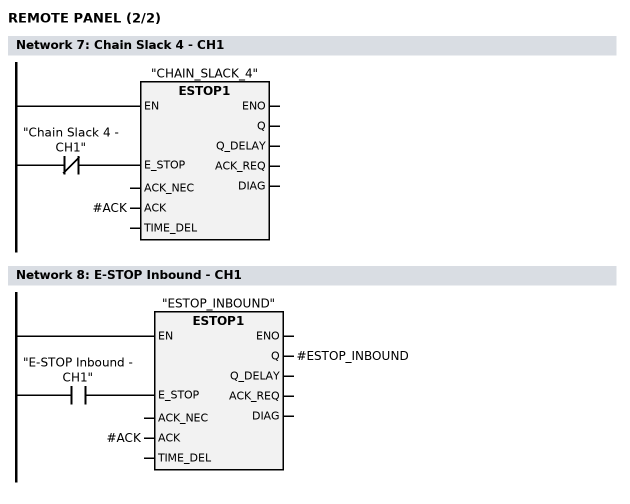
   RUNG wire#powerrail
      "CHAIN_SLACK_4".ESTOP1(E_STOP := wire#w1, ACK_NEC :=, ACK := #ACK, TIME_DEL :=, Q =>, Q_DELAY =>, ACK_REQ =>, DIAG =>)
   END_RUNG
   RUNG wire#powerrail
      I_Contact( "Chain Slack 4 - CH1" )
   END_RUNG wire#w1
   // the same network as SCL:
   "CHAIN_SLACK_4"(E_STOP := NOT "Chain Slack 4 - CH1", ACK := #ACK);   // ESTOP1
END_REGION

REGION Network 8: E-STOP Inbound - CH1
   RUNG wire#powerrail
      "ESTOP_INBOUND".ESTOP1(E_STOP := wire#w1, ACK_NEC :=, ACK := #ACK, TIME_DEL :=, Q => #ESTOP_INBOUND, Q_DELAY =>, ACK_REQ =>, DIAG =>)
   END_RUNG
   RUNG wire#powerrail
      Contact( "E-STOP Inbound - CH1" )
   END_RUNG wire#w1
   // the same network as SCL:
   "ESTOP_INBOUND"(E_STOP := "E-STOP Inbound - CH1", ACK := #ACK, Q => #ESTOP_INBOUND);   // ESTOP1
END_REGION
END_FUNCTION

FUNCTION "Mode_Change_F" : Void   // FC2, SCL
{ S7_Optimized_Access := 'TRUE' }
VERSION : 0.1
// stored: AutoNumber true, IsIECCheckEnabled false, SetENOAutomatically false, UDAEnableTagReadback false
   VAR_INPUT
      Mode : UInt;
   END_VAR
   VAR_TEMP
      i : UInt;
      j : UInt;
   END_VAR
BEGIN
   // REGION Change all devices
   //     "Control_DB".ECnv_Control.Instruction.Mode_Change := #Mode;
   //     "Control_DB".VTD_Control.Instruction.Mode_Change := #Mode;

   //     FOR #i := "Settings_DB".VTD_Settings.Lowest_Level TO "Settings_DB".VTD_Settings.Highest_Level DO
   //         "Control_DB".LCnv_Control.Cnv_Level_Control[#i].Cnv1_Control.Instruction.Mode_Change := #Mode;
   //         "Control_DB".LCnv_Control.Cnv_Level_Control[#i].Cnv2_Control.Instruction.Mode_Change := #Mode;
   //     END_FOR;
   // END_REGION
END_FUNCTION

FUNCTION_BLOCK "OPC_UA_Control_FB_1"   // FB26, SCL
{ S7_Optimized_Access := 'TRUE' }
VERSION : 0.1
// stored: AutoNumber true, IsIECCheckEnabled false, IsRetainMemResEnabled false, MemoryReserve 100, SetENOAutomatically false, UDAEnableTagReadback false
   VAR_INPUT
      OPC_Enable : Bool;
      Mode_Change : UInt;
   END_VAR
   VAR_OUTPUT
      Mode_Current : UInt;
   END_VAR
   VAR
      Source_Location_VTD { ExternalAccessible := 'False'; ExternalVisible := 'False'; ExternalWritable := 'False'} : "ID_Decoded";
      Destination_Location_VTD { ExternalAccessible := 'False'; ExternalVisible := 'False'; ExternalWritable := 'False'} : "ID_Decoded";
      Source_Location_Carousel { ExternalAccessible := 'False'; ExternalVisible := 'False'; ExternalWritable := 'False'} : "ID_Decoded";
      Destination_Location_Carousel { ExternalAccessible := 'False'; ExternalVisible := 'False'; ExternalWritable := 'False'} : "ID_Decoded";
      State_VTD : UInt;
      State_Carrousel : UInt;
   END_VAR
   VAR_TEMP
      i : UInt;
      j : UInt;
      f : UInt;
   END_VAR
BEGIN

   REGION TODO
       (*
       1. Need to confirm how the mode control is going to work, does switching the VTD to auto force all conveyors to auto as well or do we do seperate checks
       2. Need to review the shuttle interlock procedure inside the VTD function block
       *)

   END_REGION

   IF "FirstScan" THEN
       "OPC_Enable" := TRUE;
   END_IF;

   REGION Mode Control
       (*
           Mode select is done via the HMI. Might add external mode select switches.

           Mode select mask:
           0: Disabled
           1: Manual
           2: Semi-Auto
           3: Auto
           4: Teach
           5: Maintenance
       *)

       // IF #Mode_Change <> #Mode_Current THEN
       //     //Disable all devices
       //     "Mode_Change_F"(Mode := #Mode_Change);
       // END_IF;
   END_REGION

   REGION Errors VTD STATE
       IF #State_VTD > 30 AND #State_VTD < 120 THEN
           IF #Source_Location_VTD.Device_Type = 10 OR #Destination_Location_VTD.Device_Type = 10 THEN
               IF "Control_DB".LCnv_Control[#Source_Location_VTD.Level].Error
                   OR
                   "Control_DB".LCnv_Control[#Destination_Location_VTD.Level].Error THEN
                   #State_VTD := 400;
               END_IF;
           END_IF;
           IF "Control_DB".ECnv_Control.Error THEN
               #State_VTD := 400;
           END_IF;
           IF "VTD_FB_DB".I_State = 400 THEN
               #State_VTD := 400;
           END_IF;

       END_IF;
   END_REGION

   // REGION Errors CAROUSEL STATE
   //     IF #State_Carrousel > 30 AND #State_Carrousel < 120 THEN
   //         IF #Source_Location_Carousel.Device_Type = 10 OR #Destination_Location_VTD.Device_Type = 10 THEN
   //             IF "Control_DB".LCnv_Control[#Source_Location_Carousel.Level].Error
   //                 OR
   //                 "Control_DB".LCnv_Control[#Destination_Location_VTD.Level].Error THEN
   //                 #State_Carrousel := 400;
   //             END_IF;
   //         ELSIF #Source_Location_Carousel.Device_Type = 11 OR #Destination_Location_VTD.Device_Type = 11 THEN
   //             IF "Control_DB".LCnv_Control[#Source_Location_Carousel.Level].Error
   //                 OR
   //                 "Control_DB".LCnv_Control[#Destination_Location_VTD.Level].Error
   //             THEN
   //                 #State_Carrousel := 400;
   //             END_IF;
   //         END_IF;
   //         IF "Control_DB".ECnv_Control.Error THEN
   //             #State_Carrousel := 400;
   //         END_IF;
   //         IF "VTD_FB_DB".I_State = 400 THEN
   //             #State_Carrousel := 400;
   //         END_IF;

   //     END_IF;
   // END_REGION

   //Bit OPC in Error
   IF #State_VTD = 400 OR #State_Carrousel = 400 THEN
       "Error_Word_1".%X0 := TRUE;
   ELSE
       "Error_Word_1".%X0 := FALSE;
   END_IF;

   REGION OPC UA Control
       (*
       Type of task to be performed:
           1 = Move to Floor
           2 = Shuttle Transfer into VTD
           3 = Shuttle Transfer out of VTD
           4 = Transfer Pallet into VTD
           5 = Transfer Pallet out of VTD
           6 = Transfer Pallet Roller to Roller
           7 = Transfer Pallet Chain to Chain  
           8 = Transfer to pick station 
           9 = Transfer from Pick station 
           10 = Weigh Pallet
           11 = Set chain Cnv as active (lower) // no use for now
           12 = Set Roller Cnv as active (raise) // no use for now

           Need to isolate ZZ in XXYYZZ to confirm #i = ZZ

           Extract XX (first two digits)
           xx := inputNumber / 10000;

           Extract YY (middle two digits)
           yy := (inputNumber / 100) MOD 100;

           Extract ZZ (last two digits)
           zz := inputNumber MOD 100;    
       *)

       REGION VTDs and Buffer conveyors
           IF "VTD_Buffers_In_Automatic" AND #OPC_Enable THEN
               CASE #State_VTD OF
                   0:  //Pre operational state
                       #State_VTD := 10;

                   10: //Idle waiting for task
                       IF "Control_DB"."VTD_Order Table".Task_Data_Available AND "Control_DB".VTD_Control.Mode = 3 AND
                           NOT "Control_DB".VTD_Control.Running AND NOT "Control_DB"."VTD_Order Table".Movement_Ready AND "Control_DB".VTD_Control.SM_State <= 10 THEN
                               // "Control_DB".WMS_OPC_UA.Task_Data_Available := FALSE;
                               #State_VTD := 20;
                           END_IF;

                   20: //Determine the type of task
                       "ID_Decode_F"(ID := "Control_DB"."VTD_Order Table".Source_Location,
                                     ID_Decoded := #Source_Location_VTD);
                       "ID_Decode_F"(ID := "Control_DB"."VTD_Order Table".Destination_Location,
                                     ID_Decoded := #Destination_Location_VTD);

                       //VTD move to floor
                       IF "Control_DB"."VTD_Order Table".Task_Type = 1
                           AND NOT "Control_DB".VTD_Control.Running THEN
                           #State_VTD := 30;

                           //Shuttle transfer in/out of the VTD
                       ELSIF "Control_DB"."VTD_Order Table".Task_Type = 2 OR "Control_DB"."VTD_Order Table".Task_Type = 3
                       THEN
                           #State_VTD := 70;

                           //Transfer Pallet in/out of the VTD
                       ELSIF "Control_DB"."VTD_Order Table".Task_Type = 4 OR "Control_DB"."VTD_Order Table".Task_Type = 5
                       THEN
                           #State_VTD := 100;
                       END_IF;

                           //=========================== VTD Move to floor ===========================
                       30: //Set all the Move to level variables
                           "Control_DB".VTD_Control.Current_Task_Type := INT_TO_UINT("Control_DB"."VTD_Order Table".Task_Type);
                           "Control_DB".VTD_Control.Instruction.Pallet_Type := "Control_DB"."VTD_Order Table".Pallet_Type;
                           "Control_DB".VTD_Control.Instruction.Task_ID := INT_TO_UINT("Control_DB"."VTD_Order Table".Task_ID);
                           "Control_DB".VTD_Control.Instruction.Task_Metadata := "Control_DB"."VTD_Order Table".Task_Metadata;
                           "Control_DB".VTD_Control.Instruction.Move_To_Level := INT_TO_UINT(#Destination_Location_VTD.Level);
                           #State_VTD := 35;

                       35://Wait for the VTD to start its movement
                           "Control_DB"."VTD_Order Table".SM_State := "Control_DB".VTD_Control.SM_State;
                           IF "Control_DB".VTD_Control.Enabled AND "Control_DB".VTD_Control.Running THEN
                               "Control_DB"."VTD_Order Table".Movement_Ready := TRUE;
                              // "Control_DB"."VTD_Order Table".Task_Data_Available := FALSE;//
                               #State_VTD := 40;
                           END_IF;

                       40: //Wait for the VTD to complete its movement
                           "Control_DB"."VTD_Order Table".SM_State := "Control_DB".VTD_Control.SM_State;
                           IF "Control_DB".VTD_Control.SM_State = 100 THEN
                               "Control_DB"."VTD_Order Table".Movement_Request_Complete := TRUE;
                               #State_VTD := 41;
                           END_IF;

                       41: //Wait for XXs for report done
                           "IEC_Timer_0_DB_6".TON(IN := TRUE,
                                                   PT := T#2s);
                           IF "IEC_Timer_0_DB_6".Q THEN
                               #State_VTD := 45;
                           END_IF;

                       45: //Wait for the ACK before we go back to Idle
                           "Control_DB"."VTD_Order Table".SM_State := "Control_DB".VTD_Control.SM_State;
                           IF "Control_DB"."VTD_Order Table".Movement_Request_Complete_Ack THEN///////////////////////////////////////////////////////////////////
                               // "Control_DB".WMS_OPC_UA.Task_Type := 0;
                               // "Control_DB".VTD_Control.Instruction.Reset := TRUE;///////////////////////////////////////////////////////////////////
                               #State_VTD := 250;
                           END_IF;

                           //=========================== Transfer Shuttle in/out of the VTD ===========================

                       70: //Set all the shuttle interlock variables
                           "Control_DB".VTD_Control.Instruction.Task_ID := "Control_DB"."VTD_Order Table".Task_ID; //Assign task ID to WCS Task ID
                           "Control_DB".VTD_Control.Instruction.Task_Metadata := "Control_DB"."VTD_Order Table".Task_Metadata;
                           "Control_DB".VTD_Control.Instruction.Pallet_Type := "Control_DB"."VTD_Order Table".Pallet_Type;
                           "Control_DB".VTD_Control.Current_Task_Type := INT_TO_UINT("Control_DB"."VTD_Order Table".Task_Type);
                           "Control_DB".VTD_Control.Shuttle_Interlock.Shuttle_Interlock_Task_ID := INT_TO_UINT("Control_DB"."VTD_Order Table".Task_ID);
                           "Control_DB".VTD_Control.Shuttle_Interlock.Shuttle_Interlock_Task_Metadata := "Control_DB"."VTD_Order Table".Task_Metadata;
                           "Control_DB".VTD_Control.Shuttle_Interlock.Shuttle_ID := INT_TO_UINT("Control_DB"."VTD_Order Table".Shuttle_ID);
                           "Control_DB".VTD_Control.Shuttle_Interlock.Shuttle_Loaded := "Control_DB"."VTD_Order Table".Shuttle_Loaded;
                           "Control_DB".VTD_Control.Shuttle_Interlock.Shuttle_Start_Location := "Control_DB"."VTD_Order Table".Source_Location;
                           "Control_DB".VTD_Control.Shuttle_Interlock.Shuttle_Target_Location := "Control_DB"."VTD_Order Table".Destination_Location;

                           "Control_DB".VTD_Control.Shuttle_Interlock.Interlock_Request := TRUE;
                           #State_VTD := 75;

                       75: //Inform WCS that the VTD is ready to interlock
                           "Control_DB"."VTD_Order Table".SM_State := "Control_DB".VTD_Control.SM_State;
                           IF "Control_DB".VTD_Control.Shuttle_Interlock.Ready_To_Interlock THEN
                               "Control_DB"."VTD_Order Table".Movement_Ready := TRUE;
                               "Control_DB"."VTD_Order Table".Task_Data_Available := FALSE;
                               #State_VTD := 80;
                           END_IF;

                       80://Inform WCS that the interlock is complete
                           IF "Control_DB".VTD_Control.Shuttle_Interlock.Interlock_Complete THEN
                               "Control_DB".VTD_Control.Shuttle_Interlock.Interlock_Request := FALSE;
                               "Control_DB"."VTD_Order Table".Movement_Request_Complete := TRUE;
                               #State_VTD := 81;
                           END_IF;

                       81: //Wait for XXs for report done
                           "IEC_Timer_0_DB_7".TON(IN := TRUE,
                                                   PT := T#2S);
                           IF "IEC_Timer_0_DB_7".Q THEN
                               #State_VTD := 90;
                           END_IF;

                       90: //Reset VTD back to idle state
                           IF "Control_DB"."VTD_Order Table".Movement_Request_Complete_Ack THEN
                               "Control_DB".VTD_Control.Shuttle_Interlock.Interlock_Complete_Ack := TRUE;
                               #State_VTD := 250;
                           END_IF;

                           //=========================== Transfer Pallet in/out of the VTD ===========================

                       100: //Set the destination conveyor variables

                           //Assign task to receiving conveyor
                           IF #Destination_Location_VTD.Level >= "Settings_DB".VTD_Settings.Lowest_Level AND #Destination_Location_VTD.Level <= "Settings_DB".VTD_Settings.Highest_Level THEN

                               //Buffer conveyors
                               IF #Destination_Location_VTD.Device_Type = 10 AND "Control_DB".ECnv_Control.Cnv_Occupied AND
                                   NOT "Control_DB".LCnv_Control[#Destination_Location_VTD.Level].Cnv_Occupied
                               THEN
                                   "Control_DB".LCnv_Control[#Destination_Location_VTD.Level].Instruction.Task_ID := INT_TO_UINT("Control_DB"."VTD_Order Table".Task_ID);
                                   "Control_DB".LCnv_Control[#Destination_Location_VTD.Level].Instruction.Task_Metadata := "Control_DB"."VTD_Order Table".Task_Metadata;
                                   "Control_DB".LCnv_Control[#Destination_Location_VTD.Level].Current_Task_Type := INT_TO_UINT("Control_DB"."VTD_Order Table".Task_Type);
                                   "Control_DB".LCnv_Control[#Destination_Location_VTD.Level].Instruction.Transfer_From_ID := "Control_DB"."VTD_Order Table".Source_Location;
                                   "Control_DB".LCnv_Control[#Destination_Location_VTD.Level].Instruction.Transfer_To_ID := 0;

                                   //Enable the conveyor and start the transfer
                                   "Control_DB".LCnv_Control[#Destination_Location_VTD.Level].Instruction.Start_Transfer := TRUE;
                                   #State_VTD := 105;

                                  //Extractor Cnv
                               ELSIF (#Destination_Location_VTD.Device_Type = 12 AND #Source_Location_VTD.Device_Type = 10 AND NOT "Control_DB".ECnv_Control.Cnv_Occupied AND "Control_DB".LCnv_Control[#Destination_Location_VTD.Level].Cnv_Occupied)
                               THEN //FROM ECONVEYOR TO CNV1 OR CNV2
                                   "Control_DB".ECnv_Control.Instruction.Task_ID := INT_TO_UINT("Control_DB"."VTD_Order Table".Task_ID);
                                   "Control_DB".ECnv_Control.Instruction.Task_Metadata := "Control_DB"."VTD_Order Table".Task_Metadata;
                                   "Control_DB".ECnv_Control.Current_Task_Type := INT_TO_UINT("Control_DB"."VTD_Order Table".Task_Type);
                                   "Control_DB".ECnv_Control.Instruction.Transfer_From_ID := "Control_DB"."VTD_Order Table".Source_Location;
                                   "Control_DB".ECnv_Control.Instruction.Transfer_To_ID := 0;

                                   //Enable the conveyor and start the transfer
                                   "Control_DB".ECnv_Control.Instruction.Start_Transfer := TRUE;
                                   #State_VTD := 105;
                               ELSE
                                   "Error_Word_1".%X1 := TRUE; //DESTINATION CONVEYOR IS OCCUPIED
                                   #State_VTD := 400; //ERROR
                               END_IF;

                           ELSIF #Destination_Location_VTD.Level = 0 THEN
                               //Popup 2
                               IF #Destination_Location_VTD.Device_Type = 16 AND "Control_DB".ECnv_Control.Cnv_Occupied AND
                                   NOT "Control_DB".PopUp_Cnv[2].Cnv_Occupied AND "Control_DB".PopUp_Cnv[2].Inputs."Lift Down"
                               THEN//ALL GOOD
                                   "Control_DB".PopUp_Cnv[2].Instruction.Task_ID := INT_TO_UINT("Control_DB"."VTD_Order Table".Task_ID);
                                   "Control_DB".PopUp_Cnv[2].Instruction.Task_Metadata := "Control_DB"."VTD_Order Table".Task_Metadata;
                                   "Control_DB".PopUp_Cnv[2].Current_Task_Type := INT_TO_UINT("Control_DB"."VTD_Order Table".Task_Type);
                                   "Control_DB".PopUp_Cnv[2].Instruction.Transfer_From_ID := "Control_DB"."VTD_Order Table".Source_Location;
                                   "Control_DB".PopUp_Cnv[2].Instruction.Transfer_To_ID := 0;

                                   //Enable the conveyor and start the transfer
                                   "Control_DB".PopUp_Cnv[2].Instruction.Start_Transfer := TRUE;
                                   #State_VTD := 105;

                                   //Popup 2 LIFT
                               ELSIF #Destination_Location_VTD.Device_Type = 16 AND "Control_DB".ECnv_Control.Cnv_Occupied AND
                                   NOT "Control_DB".PopUp_Cnv[2].Cnv_Occupied AND NOT "Control_DB".PopUp_Cnv[2].Inputs."Lift Down"
                               THEN//NEED TO LIFT DOWN
                                   "Control_DB".PopUp_Cnv[2].Instruction.Task_ID := INT_TO_UINT("Control_DB"."VTD_Order Table".Task_ID);
                                   "Control_DB".PopUp_Cnv[2].Instruction.Task_Metadata := "Control_DB"."VTD_Order Table".Task_Metadata;
                                   "Control_DB".PopUp_Cnv[2].Current_Task_Type := INT_TO_UINT("Control_DB"."VTD_Order Table".Task_Type);
                                   "Control_DB".PopUp_Cnv[2].Instruction.Transfer_From_ID := "Control_DB"."VTD_Order Table".Source_Location;
                                   "Control_DB".PopUp_Cnv[2].Instruction.Transfer_To_ID := 0;
                                   "Control_DB".PopUp_Cnv[2].Instruction.Lift_Down := NOT "Control_DB".PopUp_Cnv[2].Running AND NOT "Control_DB".PopUp_Cnv[2].Inputs."Lift Down";
                                   IF "Control_DB".PopUp_Cnv[2].Inputs."Lift Down" THEN
                                       //Enable the conveyor and start the transfer
                                       "Control_DB".PopUp_Cnv[2].Instruction.Start_Transfer := TRUE;
                                       #State_VTD := 105;
                                   END_IF;

                                   //Extractor Cnv
                               ELSIF (#Destination_Location_VTD.Device_Type = 12 AND #Source_Location_VTD.Device_Type = 16 AND NOT "Control_DB".ECnv_Control.Cnv_Occupied AND "Control_DB".PopUp_Cnv[2].Cnv_Occupied)
                               THEN //FROM ECONVEYOR TO CNV1 OR CNV2
                                   "Control_DB".ECnv_Control.Instruction.Task_ID := INT_TO_UINT("Control_DB"."VTD_Order Table".Task_ID);
                                   "Control_DB".ECnv_Control.Instruction.Task_Metadata := "Control_DB"."VTD_Order Table".Task_Metadata;
                                   "Control_DB".ECnv_Control.Current_Task_Type := INT_TO_UINT("Control_DB"."VTD_Order Table".Task_Type);
                                   "Control_DB".ECnv_Control.Instruction.Transfer_From_ID := "Control_DB"."VTD_Order Table".Source_Location;
                                   "Control_DB".ECnv_Control.Instruction.Transfer_To_ID := 0;

                                   //Enable the conveyor and start the transfer
                                   "Control_DB".ECnv_Control.Instruction.Start_Transfer := TRUE;
                                   #State_VTD := 105;
                               ELSE
                                   "Error_Word_1".%X1 := TRUE; //DESTINATION CONVEYOR IS OCCUPIED
                                   #State_VTD := 400; //ERROR
                               END_IF;
                           ELSE
                               ; //Error: the destination location is not possible
                               #State_VTD := 400;
                           END_IF;

                       105:  //Set the source conveyor variables

                           //Assign task to sending conveyor
                           IF #Source_Location_VTD.Level >= "Settings_DB".VTD_Settings.Lowest_Level AND #Source_Location_VTD.Level <= "Settings_DB".VTD_Settings.Highest_Level THEN

                               //Cnv_Front_of_VTD
                               IF #Source_Location_VTD.Device_Type = 10 AND NOT "Control_DB".ECnv_Control.Cnv_Occupied AND "Control_DB".LCnv_Control[#Source_Location_VTD.Level].Cnv_Occupied THEN //FROM CONV1 TO ECONVEYOR
                                   "Control_DB".LCnv_Control[#Source_Location_VTD.Level].Instruction.Task_ID := INT_TO_UINT("Control_DB"."VTD_Order Table".Task_ID);
                                   "Control_DB".LCnv_Control[#Source_Location_VTD.Level].Instruction.Task_Metadata := "Control_DB"."VTD_Order Table".Task_Metadata;
                                   "Control_DB".LCnv_Control[#Source_Location_VTD.Level].Current_Task_Type := INT_TO_UINT("Control_DB"."VTD_Order Table".Task_Type);
                                   "Control_DB".LCnv_Control[#Source_Location_VTD.Level].Instruction.Transfer_To_ID := "Control_DB"."VTD_Order Table".Destination_Location;
                                   "Control_DB".LCnv_Control[#Source_Location_VTD.Level].Instruction.Transfer_From_ID := 0;

                                   //Enable the conveyor and start the transfer
                                   "Control_DB".LCnv_Control[#Source_Location_VTD.Level].Instruction.Start_Transfer := TRUE;
                                   #State_VTD := 110;

                                   //Extractor Cnv
                               ELSIF (#Source_Location_VTD.Device_Type = 12 AND #Destination_Location_VTD.Device_Type = 10 AND "Control_DB".ECnv_Control.Cnv_Occupied AND NOT "Control_DB".LCnv_Control[#Source_Location_VTD.Level].Cnv_Occupied)
                               THEN //FROM ECONVEYOR TO CNV1 OR CNV2
                                   "Control_DB".ECnv_Control.Instruction.Task_ID := INT_TO_UINT("Control_DB"."VTD_Order Table".Task_ID);
                                   "Control_DB".ECnv_Control.Instruction.Task_Metadata := "Control_DB"."VTD_Order Table".Task_Metadata;
                                   "Control_DB".ECnv_Control.Current_Task_Type := INT_TO_UINT("Control_DB"."VTD_Order Table".Task_Type);
                                   "Control_DB".ECnv_Control.Instruction.Transfer_To_ID := "Control_DB"."VTD_Order Table".Destination_Location;
                                   "Control_DB".ECnv_Control.Instruction.Transfer_From_ID := 0;

                                   //Enable the conveyor and start the transfer
                                   "Control_DB".ECnv_Control.Instruction.Start_Transfer := TRUE;
                                   #State_VTD := 110;
                               ELSE
                                   "Error_Word_1".%X1 := TRUE; //DESTINATION CONVEYOR IS OCCUPIED
                                   #State_VTD := 400; //ERROR
                               END_IF;

                           ELSIF #Source_Location_VTD.Level = 0 THEN
                               //PopUp conveyor 2   
                               IF #Source_Location_VTD.Device_Type = 16 AND NOT "Control_DB".ECnv_Control.Cnv_Occupied AND
                                   "Control_DB".PopUp_Cnv[2].Cnv_Occupied AND "Control_DB".PopUp_Cnv[2].Inputs."Lift Down" THEN //FROM CONV2 TO ECONVEYOR
                                   "Control_DB".PopUp_Cnv[2].Instruction.Task_ID := INT_TO_UINT("Control_DB"."VTD_Order Table".Task_ID);
                                   "Control_DB".PopUp_Cnv[2].Instruction.Task_Metadata := "Control_DB"."VTD_Order Table".Task_Metadata;
                                   "Control_DB".PopUp_Cnv[2].Current_Task_Type := INT_TO_UINT("Control_DB"."VTD_Order Table".Task_Type);
                                   "Control_DB".PopUp_Cnv[2].Instruction.Transfer_To_ID := "Control_DB"."VTD_Order Table".Destination_Location;
                                   "Control_DB".PopUp_Cnv[2].Instruction.Transfer_From_ID := 0;

                                   //Enable the conveyor and start the transfer
                                   "Control_DB".PopUp_Cnv[2].Instruction.Start_Transfer := TRUE;
                                   #State_VTD := 110;

                                   //Popup 2 LIFT
                               ELSIF #Source_Location_VTD.Device_Type = 16 AND NOT "Control_DB".ECnv_Control.Cnv_Occupied AND
                                   "Control_DB".PopUp_Cnv[2].Cnv_Occupied AND NOT "Control_DB".PopUp_Cnv[2].Inputs."Lift Down"
                               THEN//NEED TO LIFT DOWN
                                   "Control_DB".PopUp_Cnv[2].Instruction.Task_ID := INT_TO_UINT("Control_DB"."VTD_Order Table".Task_ID);
                                   "Control_DB".PopUp_Cnv[2].Instruction.Task_Metadata := "Control_DB"."VTD_Order Table".Task_Metadata;
                                   "Control_DB".PopUp_Cnv[2].Current_Task_Type := INT_TO_UINT("Control_DB"."VTD_Order Table".Task_Type);
                                   "Control_DB".PopUp_Cnv[2].Instruction.Transfer_From_ID := 0;
                                   "Control_DB".PopUp_Cnv[2].Instruction.Transfer_To_ID := "Control_DB"."VTD_Order Table".Destination_Location;
                                   "Control_DB".PopUp_Cnv[2].Instruction.Lift_Down := NOT "Control_DB".PopUp_Cnv[2].Running AND NOT "Control_DB".PopUp_Cnv[2].Inputs."Lift Down";
                                   IF "Control_DB".PopUp_Cnv[2].Inputs."Lift Down" THEN
                                       //Enable the conveyor and start the transfer
                                       "Control_DB".PopUp_Cnv[2].Instruction.Start_Transfer := TRUE;
                                       #State_VTD := 110;
                                   END_IF;

                                   //Extractor Cnv
                               ELSIF (#Source_Location_VTD.Device_Type = 12 AND #Destination_Location_VTD.Device_Type = 16 AND "Control_DB".ECnv_Control.Cnv_Occupied AND NOT "Control_DB".PopUp_Cnv[2].Cnv_Occupied)
                               THEN //FROM ECONVEYOR TO CNV1 OR CNV2
                                   "Control_DB".ECnv_Control.Instruction.Task_ID := INT_TO_UINT("Control_DB"."VTD_Order Table".Task_ID);
                                   "Control_DB".ECnv_Control.Instruction.Task_Metadata := "Control_DB"."VTD_Order Table".Task_Metadata;
                                   "Control_DB".ECnv_Control.Current_Task_Type := INT_TO_UINT("Control_DB"."VTD_Order Table".Task_Type);
                                   "Control_DB".ECnv_Control.Instruction.Transfer_To_ID := "Control_DB"."VTD_Order Table".Destination_Location;
                                   "Control_DB".ECnv_Control.Instruction.Transfer_From_ID := 0;

                                   //Enable the conveyor and start the transfer
                                   "Control_DB".ECnv_Control.Instruction.Start_Transfer := TRUE;
                                   #State_VTD := 110;
                               END_IF;
                           ELSE
                               ; //Error: the destination location is not possible
                               #State_VTD := 400;
                           END_IF;

                       110: //Start the transfer
                           "Control_DB"."VTD_Order Table".SM_State := "Control_DB".ECnv_Control.SM_State;
                           IF "Control_DB".ECnv_Control.Enabled AND "Control_DB".ECnv_Control.Running THEN
                               "Control_DB"."VTD_Order Table".Movement_Ready := TRUE;
                               "Control_DB"."VTD_Order Table".Task_Data_Available := FALSE;
                               #State_VTD := 115;
                           END_IF;

                       115: //Wait for the transfer to complete
                           "Control_DB"."VTD_Order Table".SM_State := "Control_DB".ECnv_Control.SM_State;
                           IF "Control_DB".ECnv_Control.Done THEN
                               "Control_DB".ECnv_Control.Instruction.Start_Transfer := FALSE;
                               "Control_DB".LCnv_Control[1].Instruction.Start_Transfer := FALSE;
                               "Control_DB".LCnv_Control[2].Instruction.Start_Transfer := FALSE;
                               "Control_DB".LCnv_Control[3].Instruction.Start_Transfer := FALSE;
                               "Control_DB".PopUp_Cnv[2].Instruction.Start_Transfer := FALSE;
                               "Control_DB"."VTD_Order Table".Movement_Request_Complete := TRUE;
                               #State_VTD := 116;
                           END_IF;

                       116: //Wait for XXs for report done
                           "IEC_Timer_0_DB_5".TON(IN := TRUE,
                                                   PT := T#2S);
                           IF "IEC_Timer_0_DB_5".Q THEN
                               #State_VTD := 120;
                           END_IF;

                       120: //Wait for the ACK before we go back to Idle
                           "Control_DB"."VTD_Order Table".SM_State := "Control_DB".ECnv_Control.SM_State;
                           IF "Control_DB"."VTD_Order Table".Movement_Request_Complete_Ack THEN
                               // "Control_DB".ECnv_Control.Instruction.Reset := TRUE;
                               #State_VTD := 250;
                           END_IF;

                           //=========================== Reset and Error States ===========================
                       250: //Reset all variable and return to idle

                           //Reset the OPC control variables
                           "Control_DB"."VTD_Order Table".SM_State := 0;
                           "Control_DB"."VTD_Order Table".Movement_Ready := FALSE;
                           "Control_DB"."VTD_Order Table".Movement_Request_Complete := FALSE;
                           "Control_DB"."VTD_Order Table".Movement_Request_Complete_Ack := FALSE;
                           "Control_DB"."VTD_Order Table".Task_Metadata := '';
                           "IEC_Timer_0_DB_5".TON(IN := FALSE,
                                                  PT := T#0S);
                           "IEC_Timer_0_DB_6".TON(IN := FALSE,
                                                  PT := T#0S);
                           "IEC_Timer_0_DB_7".TON(IN := FALSE,
                                                  PT := T#0S);

                           // Reset Order table VTD variables
                           "Control_DB"."VTD_Order Table".Task_Type := 0;
                           "Control_DB"."VTD_Order Table".Pallet_Type:='C';
                           "Control_DB"."VTD_Order Table".Task_ID:= 0;
                           "Control_DB"."VTD_Order Table".Task_Metadata:='';
                           "Control_DB"."VTD_Order Table".Source_Location := 0;
                           "Control_DB"."VTD_Order Table".Destination_Location := 0;
                           #Destination_Location_VTD.Level:=0;
                           #Source_Location_VTD.Level := 0;
                           "Control_DB"."VTD_Order Table".Shuttle_ID := 0;
                           "Control_DB"."VTD_Order Table".Shuttle_Loaded := FALSE;


                           //Reset VTD variables
                           "Control_DB".VTD_Control.Instruction.Reset := FALSE;
                           "Control_DB".VTD_Control.Instruction.Pallet_Type := 0;
                           "Control_DB".VTD_Control.Instruction.Task_ID := 0;
                           "Control_DB".VTD_Control.Instruction.Task_Metadata := '';
                           "Control_DB".VTD_Control.Instruction.Move_To_Level := 99;
                           "Control_DB".VTD_Control.Current_Task_Type := 0;

                           //Reset Shuttle interlock
                           "Control_DB".VTD_Control.Shuttle_Interlock.Interlock_Request := FALSE;
                           "Control_DB".VTD_Control.Shuttle_Interlock.Shuttle_Start_Location := 0;
                           "Control_DB".VTD_Control.Shuttle_Interlock.Shuttle_Target_Location := 0;
                           "Control_DB".VTD_Control.Shuttle_Interlock.Shuttle_Loaded := 0;
                           "Control_DB".VTD_Control.Shuttle_Interlock.Shuttle_ID := 0;
                           "Control_DB".VTD_Control.Shuttle_Interlock.Shuttle_Interlock_Task_ID := 0;
                           "Control_DB".VTD_Control.Shuttle_Interlock.Shuttle_Interlock_Task_Metadata := '';
                           "Control_DB".VTD_Control.Shuttle_Interlock.Interlock_Complete_Ack := FALSE;

                           //Reset conveyor variables
                           "Control_DB".ECnv_Control.Instruction.Reset := FALSE;
                           // "Control_DB".ECnv_Control.Instruction.Enable := FALSE;
                           "Control_DB".ECnv_Control.Instruction.Start_Transfer := FALSE;
                           "Control_DB".ECnv_Control.Instruction.Task_ID := 0;
                           "Control_DB".ECnv_Control.Instruction.Task_Metadata := '';
                           "Control_DB".ECnv_Control.Current_Task_Type := 0;
                           "Control_DB".ECnv_Control.Instruction.Transfer_From_ID := 0;
                           "Control_DB".ECnv_Control.Instruction.Transfer_To_ID := 0;

                           FOR #i := "Settings_DB".VTD_Settings.Lowest_Level TO "Settings_DB".VTD_Settings.Highest_Level DO
                               "Control_DB".LCnv_Control[#i].Instruction.Reset := FALSE;
                               "Control_DB".LCnv_Control[#i].Instruction.Start_Transfer := FALSE;
                               "Control_DB".LCnv_Control[#i].Instruction.Task_ID := 0;
                               "Control_DB".LCnv_Control[#i].Instruction.Task_Metadata := '';
                               "Control_DB".LCnv_Control[#i].Current_Task_Type := 0;
                               "Control_DB".LCnv_Control[#i].Instruction.Transfer_From_ID := 0;
                               "Control_DB".LCnv_Control[#i].Instruction.Transfer_To_ID := 0;

                               "Control_DB".LCnv_Control[#i].Instruction.Reset := FALSE;
                               "Control_DB".LCnv_Control[#i].Instruction.Start_Transfer := FALSE;
                               "Control_DB".LCnv_Control[#i].Instruction.Task_ID := 0;
                               "Control_DB".LCnv_Control[#i].Instruction.Task_Metadata := '';
                               "Control_DB".LCnv_Control[#i].Current_Task_Type := 0;
                               "Control_DB".LCnv_Control[#i].Instruction.Transfer_From_ID := 0;
                               "Control_DB".LCnv_Control[#i].Instruction.Transfer_To_ID := 0;
                           END_FOR;

                           "Control_DB".PopUp_Cnv[2].Instruction.Start_Transfer := FALSE;
                           "Control_DB".PopUp_Cnv[2].Instruction.Task_ID := 0;
                           "Control_DB".PopUp_Cnv[2].Instruction.Task_Metadata := '';
                           "Control_DB".PopUp_Cnv[2].Current_Task_Type := 0;
                           "Control_DB".PopUp_Cnv[2].Instruction.Transfer_From_ID := 0;
                           "Control_DB".PopUp_Cnv[2].Instruction.Transfer_To_ID := 0;

                           "Error_Word_1".%X1 := FALSE;

                           #State_VTD := 0;

                       400:// Error state
                           "Control_DB".VTD_Control.Shuttle_Interlock.Interlock_Request := FALSE;
                           "Control_DB".VTD_Control.Shuttle_Interlock.Interlock_Complete_Ack := FALSE;
                           "Control_DB"."VTD_Order Table".Task_Metadata := '';
                           // Reset Order table VTD variables
                           "Control_DB"."VTD_Order Table".Task_Type := 0;
                           "Control_DB"."VTD_Order Table".Pallet_Type := 'C';
                           "Control_DB"."VTD_Order Table".Task_ID := 0;
                           "Control_DB"."VTD_Order Table".Task_Metadata := '';
                           "Control_DB"."VTD_Order Table".Source_Location := 0;
                           "Control_DB"."VTD_Order Table".Destination_Location := 0;
                           #Destination_Location_VTD.Level := 0;
                           #Source_Location_VTD.Level := 0;
                           "Control_DB"."VTD_Order Table".Shuttle_ID := 0;
                           "Control_DB"."VTD_Order Table".Shuttle_Loaded := FALSE;

                           IF "Control_DB".VTD_Control.Instruction.Reset
                           THEN
                               #State_VTD := 250;
                           END_IF;

                           ELSE
                               ;
                       END_CASE;
                   ELSIF "VTD_Buffers_In_Automatic" AND NOT #OPC_Enable THEN
                       "Control_DB"."VTD_Order Table".Task_Metadata := '';
                       //Reset all variable and return to idle

                       //Reset the OPC control variables
                       "Control_DB"."VTD_Order Table".SM_State := 0;
                       "Control_DB"."VTD_Order Table".Movement_Ready := FALSE;
                       "Control_DB"."VTD_Order Table".Movement_Request_Complete := FALSE;

                       // Reset Order table VTD variables
                       "Control_DB"."VTD_Order Table".Task_Type := 0;
                       "Control_DB"."VTD_Order Table".Pallet_Type := 'C';
                       "Control_DB"."VTD_Order Table".Task_ID := 0;
                       "Control_DB"."VTD_Order Table".Task_Metadata := '';
                       "Control_DB"."VTD_Order Table".Source_Location := 0;
                       "Control_DB"."VTD_Order Table".Destination_Location := 0;
                       #Destination_Location_VTD.Level := 0;
                       #Source_Location_VTD.Level := 0;
                       "Control_DB"."VTD_Order Table".Shuttle_ID := 0;
                       "Control_DB"."VTD_Order Table".Shuttle_Loaded := FALSE;

                       //Reset VTD variables
                       "Control_DB".VTD_Control.Instruction.Reset := FALSE;
                       "Control_DB".VTD_Control.Instruction.Pallet_Type := 0;
                       "Control_DB".VTD_Control.Instruction.Task_ID := 0;
                       "Control_DB".VTD_Control.Instruction.Task_Metadata := '';//
                       "Control_DB".ECnv_Control.Current_Task_Type := 0;
                       "Control_DB".VTD_Control.Instruction.Move_To_Level := 99;
                       "Control_DB".VTD_Control.Current_Task_Type := 0;

                       //Reset Shuttle interlock
                       "Control_DB".VTD_Control.Shuttle_Interlock.Interlock_Request := FALSE;
                       "Control_DB".VTD_Control.Shuttle_Interlock.Shuttle_Start_Location := 0;
                       "Control_DB".VTD_Control.Shuttle_Interlock.Shuttle_Target_Location := 0;
                       "Control_DB".VTD_Control.Shuttle_Interlock.Shuttle_Loaded := 0;
                       "Control_DB".VTD_Control.Shuttle_Interlock.Shuttle_ID := 0;
                       "Control_DB".VTD_Control.Shuttle_Interlock.Shuttle_Interlock_Task_ID := 0;
                       "Control_DB".VTD_Control.Shuttle_Interlock.Shuttle_Interlock_Task_Metadata := '';//

                       //Reset conveyor variables
                       "Control_DB".ECnv_Control.Instruction.Reset := FALSE;
                       // "Control_DB".ECnv_Control.Instruction.Enable := FALSE;
                       "Control_DB".ECnv_Control.Instruction.Start_Transfer := FALSE;
                       "Control_DB".ECnv_Control.Instruction.Task_ID := 0;
                       "Control_DB".ECnv_Control.Instruction.Task_Metadata := '';//
                       "Control_DB".ECnv_Control.Instruction.Transfer_From_ID := 0;
                       "Control_DB".ECnv_Control.Instruction.Transfer_To_ID := 0;

                       FOR #i := "Settings_DB".VTD_Settings.Lowest_Level TO "Settings_DB".VTD_Settings.Highest_Level DO
                           "Control_DB".LCnv_Control[#i].Instruction.Reset := FALSE;
                           "Control_DB".LCnv_Control[#i].Instruction.Start_Transfer := FALSE;
                           "Control_DB".LCnv_Control[#i].Instruction.Task_ID := 0;
                           "Control_DB".LCnv_Control[#i].Instruction.Task_Metadata := '';
                           "Control_DB".LCnv_Control[#i].Current_Task_Type := 0;
                           "Control_DB".LCnv_Control[#i].Instruction.Transfer_From_ID := 0;
                           "Control_DB".LCnv_Control[#i].Instruction.Transfer_To_ID := 0;

                           "Control_DB".LCnv_Control[#i].Instruction.Reset := FALSE;
                           "Control_DB".LCnv_Control[#i].Instruction.Start_Transfer := FALSE;
                           "Control_DB".LCnv_Control[#i].Instruction.Task_ID := 0;
                           "Control_DB".LCnv_Control[#i].Instruction.Task_Metadata := '';
                           "Control_DB".LCnv_Control[#i].Current_Task_Type := 0;
                           "Control_DB".LCnv_Control[#i].Instruction.Transfer_From_ID := 0;
                           "Control_DB".LCnv_Control[#i].Instruction.Transfer_To_ID := 0;
                       END_FOR;
                   END_IF;
               END_REGION

       REGION Carrousel
           IF "Carrousel_In_Automatic" AND #OPC_Enable THEN
               CASE #State_Carrousel OF
                   0:  //Pre operational state
                       #State_Carrousel := 10;

                   10: //Idle waiting for task
                       IF "Control_DB"."Carrousel_Order Table".Task_Data_Available THEN
                           #State_Carrousel := 20;
                       END_IF;

                   20: //Determine the type of task
                       "ID_Decode_F"(ID := "Control_DB"."Carrousel_Order Table".Source_Location,
                                     ID_Decoded := #Source_Location_Carousel);
                       "ID_Decode_F"(ID := "Control_DB"."Carrousel_Order Table".Destination_Location,
                                     ID_Decoded := #Destination_Location_Carousel);

                               // Transfer Pallet Roller to Roller  
                       IF "Control_DB"."Carrousel_Order Table".Task_Type = 6 OR "Control_DB"."Carrousel_Order Table".Task_Type = 16 OR "Control_DB"."Carrousel_Order Table".Task_Type = 14 THEN
                               #State_Carrousel := 30;

                               // Transfer Pallet Chain to Chain
                           ELSIF "Control_DB"."Carrousel_Order Table".Task_Type = 7 THEN
                               #State_Carrousel := 80;

                               // Transfer to pick station (From Pop Conveyor 4)
                           ELSIF "Control_DB"."Carrousel_Order Table".Task_Type = 8 THEN
                               #State_Carrousel := 130;

                               // Transfer from Pick station (To Pop Conveyor 1)
                           ELSIF "Control_DB"."Carrousel_Order Table".Task_Type = 9 THEN
                               #State_Carrousel := 180;

                               // Start weigh measurement (Weigh Station)
                           ELSIF "Control_DB"."Carrousel_Order Table".Task_Type = 10 THEN
                               #State_Carrousel := 230;

                           END_IF;

                           //=========================== Transfer Pallet Roller to Roller  ===========================

                       30: //Check which conveyor
                               //Inbound conveyor to popup conveyor 1
                           IF #Source_Location_Carousel.Device_Type = 13 AND #Destination_Location_Carousel.Device_Type = 15 AND "Control_DB".Inbound_Cnv.Cnv_Occupied AND
                               NOT "Control_DB".PopUp_Cnv[1].Cnv_Occupied AND "Control_DB".PopUp_Cnv[1].Inputs."Lift Up"
                           THEN //All good
                               #State_Carrousel := 50;// Roller Transfer
                           ELSIF #Source_Location_Carousel.Device_Type = 13 AND #Destination_Location_Carousel.Device_Type = 15 AND "Control_DB".Inbound_Cnv.Cnv_Occupied AND
                               NOT "Control_DB".PopUp_Cnv[1].Cnv_Occupied AND NOT "Control_DB".PopUp_Cnv[1].Inputs."Lift Up"
                           THEN //Lift
                               #State_Carrousel := 40;// Lift pop up 1 

                               //Pop conveyor 1 to popup conveyor 2    
                           ELSIF #Source_Location_Carousel.Device_Type = 15 AND #Destination_Location_Carousel.Device_Type = 16 AND "Control_DB".PopUp_Cnv[1].Cnv_Occupied AND
                               NOT "Control_DB".PopUp_Cnv[2].Cnv_Occupied AND "Control_DB".PopUp_Cnv[1].Inputs."Lift Up" AND "Control_DB".PopUp_Cnv[2].Inputs."Lift Up"
                           THEN //All good
                               #State_Carrousel := 50;// Roller Transfer
                           ELSIF #Source_Location_Carousel.Device_Type = 15 AND #Destination_Location_Carousel.Device_Type = 16 AND "Control_DB".PopUp_Cnv[1].Cnv_Occupied AND
                               NOT "Control_DB".PopUp_Cnv[2].Cnv_Occupied AND (NOT "Control_DB".PopUp_Cnv[1].Inputs."Lift Up" OR NOT "Control_DB".PopUp_Cnv[2].Inputs."Lift Up")
                           THEN //Lift
                               #State_Carrousel := 40;// Lift pop up 1 OR 2

                               //Pop conveyor 3 to popup conveyor 4    
                           ELSIF #Source_Location_Carousel.Device_Type = 17 AND #Destination_Location_Carousel.Device_Type = 18 AND "Control_DB".PopUp_Cnv[3].Cnv_Occupied AND
                               NOT "Control_DB".PopUp_Cnv[4].Cnv_Occupied AND "Control_DB".PopUp_Cnv[3].Inputs."Lift Up" AND "Control_DB".PopUp_Cnv[4].Inputs."Lift Up"
                           THEN //All good
                               #State_Carrousel := 50;// Roller Transfer
                           ELSIF #Source_Location_Carousel.Device_Type = 17 AND #Destination_Location_Carousel.Device_Type = 18 AND "Control_DB".PopUp_Cnv[3].Cnv_Occupied AND
                               NOT "Control_DB".PopUp_Cnv[4].Cnv_Occupied AND (NOT "Control_DB".PopUp_Cnv[3].Inputs."Lift Up" OR NOT "Control_DB".PopUp_Cnv[4].Inputs."Lift Up")
                           THEN //Lift
                               #State_Carrousel := 40;// Lift pop up 3 OR 4

                               //Pop conveyor 4 to Outbound conveyor
                           ELSIF #Source_Location_Carousel.Device_Type = 18 AND #Destination_Location_Carousel.Device_Type = 14 AND "Control_DB".PopUp_Cnv[4].Cnv_Occupied AND
                               NOT "Control_DB".Outbound_Cnv.Cnv_Occupied AND "Control_DB".PopUp_Cnv[4].Inputs."Lift Up"
                           THEN //All good
                               #State_Carrousel := 50;// Roller Transfer
                           ELSIF #Source_Location_Carousel.Device_Type = 18 AND #Destination_Location_Carousel.Device_Type = 14 AND "Control_DB".PopUp_Cnv[4].Cnv_Occupied AND
                               NOT "Control_DB".Outbound_Cnv.Cnv_Occupied AND NOT "Control_DB".PopUp_Cnv[4].Inputs."Lift Up"
                           THEN //Lift
                               #State_Carrousel := 40;// Lift pop up 4
                           ELSE
                               ; //Error: the destination location is not possible
                               #State_Carrousel := 400;
                           END_IF;

                       40:  //Lift PopUps
                           //INBOUND CONVEYOR TO POPUP 1
                           IF #Source_Location_Carousel.Device_Type = 13 AND #Destination_Location_Carousel.Device_Type = 15 THEN
                               "Control_DB".PopUp_Cnv[1].Instruction.Lift_Up := NOT "Control_DB".PopUp_Cnv[1].Running AND NOT "Control_DB".PopUp_Cnv[1].Inputs."Lift Up";
                               IF "Control_DB".PopUp_Cnv[1].Inputs."Lift Up" THEN
                                   "Control_DB".PopUp_Cnv[1].Instruction.Lift_Up := FALSE;
                                   #State_Carrousel := 50;
                               END_IF;

                               //POPUP 1 TO 2
                           ELSIF #Source_Location_Carousel.Device_Type = 15 OR #Destination_Location_Carousel.Device_Type = 16 THEN
                               "Control_DB".PopUp_Cnv[1].Instruction.Lift_Up := NOT "Control_DB".PopUp_Cnv[1].Running AND NOT "Control_DB".PopUp_Cnv[1].Inputs."Lift Up";
                               "Control_DB".PopUp_Cnv[2].Instruction.Lift_Up := NOT "Control_DB".PopUp_Cnv[2].Running AND NOT "Control_DB".PopUp_Cnv[2].Inputs."Lift Up";
                               IF "Control_DB".PopUp_Cnv[2].Inputs."Lift Up" AND "Control_DB".PopUp_Cnv[1].Inputs."Lift Up" THEN
                                   "Control_DB".PopUp_Cnv[1].Instruction.Lift_Up := FALSE;
                                   "Control_DB".PopUp_Cnv[2].Instruction.Lift_Up := FALSE;
                                   #State_Carrousel := 50;
                               END_IF;

                               //POPUP 3 TO 4
                           ELSIF #Source_Location_Carousel.Device_Type = 17 OR #Destination_Location_Carousel.Device_Type = 18 THEN
                               "Control_DB".PopUp_Cnv[3].Instruction.Lift_Up := NOT "Control_DB".PopUp_Cnv[3].Running AND NOT "Control_DB".PopUp_Cnv[3].Inputs."Lift Up";
                               "Control_DB".PopUp_Cnv[4].Instruction.Lift_Up := NOT "Control_DB".PopUp_Cnv[4].Running AND NOT "Control_DB".PopUp_Cnv[4].Inputs."Lift Up";
                               IF "Control_DB".PopUp_Cnv[3].Inputs."Lift Up" AND "Control_DB".PopUp_Cnv[4].Inputs."Lift Up" THEN
                                   #State_Carrousel := 50;
                               END_IF;

                               //POPUP 4 TO OUTBOUND CONVEYOR
                           ELSIF #Source_Location_Carousel.Device_Type = 18 OR #Destination_Location_Carousel.Device_Type = 14 THEN
                               "Control_DB".PopUp_Cnv[4].Instruction.Lift_Up := NOT "Control_DB".PopUp_Cnv[4].Running AND NOT "Control_DB".PopUp_Cnv[4].Inputs."Lift Up";
                               IF "Control_DB".PopUp_Cnv[4].Inputs."Lift Up" THEN
                                   #State_Carrousel := 50;
                               END_IF;
                           END_IF;

                       50: //Start the transfer
                           //Inbound to popup 1 conveyors
                           IF #Source_Location_Carousel.Device_Type = 13 AND #Destination_Location_Carousel.Device_Type = 15 THEN
                               "Control_DB"."Carrousel_Order Table".SM_State := "Control_DB".PopUp_Cnv[1].SM_State;//Current machine state
                               "Control_DB".PopUp_Cnv[1].Instruction.Start_Transfer := NOT "Control_DB".PopUp_Cnv[1].Running AND "Control_DB".Inbound_Cnv.SM_State = 30;
                               "Control_DB".Inbound_Cnv.Instruction.Start_Transfer := NOT "Control_DB".Inbound_Cnv.Running ;
                               IF "Control_DB".PopUp_Cnv[1].Running AND "Control_DB".Inbound_Cnv.Running THEN
                                   "Control_DB"."Carrousel_Order Table".Movement_Ready := TRUE;
                                  // "Control_DB"."Carrousel_Order Table".Task_Data_Available := FALSE;
                                   #State_Carrousel := 60;
                               END_IF;
                           END_IF;

                           //Popup 1 TO Popup 2 conveyors
                           IF #Source_Location_Carousel.Device_Type = 15 AND #Destination_Location_Carousel.Device_Type = 16 THEN
                               "Control_DB".PopUp_Cnv[2].Instruction.Transfer_From_ID := "Settings_DB".PopUp_Cnv_Settings[1].ID;
                               "Control_DB"."Carrousel_Order Table".SM_State := "Control_DB".PopUp_Cnv[2].SM_State;//Current machine state
                               "Control_DB".PopUp_Cnv[2].Instruction.Start_Transfer := NOT "Control_DB".PopUp_Cnv[2].Running;
                               "Control_DB".PopUp_Cnv[1].Instruction.Start_Transfer := NOT "Control_DB".PopUp_Cnv[1].Running;
                               IF "Control_DB".PopUp_Cnv[2].Running AND "Control_DB".PopUp_Cnv[1].Running THEN
                                   "Control_DB"."Carrousel_Order Table".Movement_Ready := TRUE;
                                  // "Control_DB"."Carrousel_Order Table".Task_Data_Available := FALSE;
                                   #State_Carrousel := 60;
                               END_IF;
                           END_IF;

                           //Popup 3 TO Popup 4 conveyors
                           IF #Source_Location_Carousel.Device_Type = 17 AND #Destination_Location_Carousel.Device_Type = 18 THEN
                               "Control_DB"."Carrousel_Order Table".SM_State := "Control_DB".PopUp_Cnv[4].SM_State;//Current machine state
                               "Control_DB".PopUp_Cnv[4].Instruction.Start_Transfer := NOT "Control_DB".PopUp_Cnv[4].Running;
                               "Control_DB".PopUp_Cnv[3].Instruction.Start_Transfer := NOT "Control_DB".PopUp_Cnv[3].Running;
                               IF "Control_DB".PopUp_Cnv[4].Running AND "Control_DB".PopUp_Cnv[3].Running THEN
                                   "Control_DB"."Carrousel_Order Table".Movement_Ready := TRUE;
                                   "Control_DB"."Carrousel_Order Table".Task_Data_Available := FALSE;
                                   #State_Carrousel := 60;
                               END_IF;
                           END_IF;

                           //Popup 4 TO Outbound conveyors
                           IF #Source_Location_Carousel.Device_Type = 18 AND #Destination_Location_Carousel.Device_Type = 14 THEN
                               "Control_DB"."Carrousel_Order Table".SM_State := "Control_DB".Outbound_Cnv.SM_State;//Current machine state
                               "Control_DB".Outbound_Cnv.Instruction.Start_Transfer := NOT "Control_DB".Outbound_Cnv.Running;
                               "Control_DB".PopUp_Cnv[4].Instruction.Start_Transfer := NOT "Control_DB".PopUp_Cnv[4].Running;
                               IF "Control_DB".Outbound_Cnv.Running AND "Control_DB".PopUp_Cnv[4].Running THEN
                                   "Control_DB"."Carrousel_Order Table".Movement_Ready := TRUE;
                                   //"Control_DB"."Carrousel_Order Table".Task_Data_Available := FALSE;
                                   #State_Carrousel := 60;
                               END_IF;
                           END_IF;

                       60: //Wait for the transfer to complete
                           //Inbound to popup 1 conveyors
                           IF #Source_Location_Carousel.Device_Type = 13 AND #Destination_Location_Carousel.Device_Type = 15 AND
                               "Control_DB".PopUp_Cnv[1].Done AND "Control_DB".Inbound_Cnv.Done
                           THEN
                               "Control_DB"."Carrousel_Order Table".SM_State := "Control_DB".PopUp_Cnv[1].SM_State;
                               "Control_DB"."Carrousel_Order Table".Movement_Request_Complete := TRUE;
                               #State_Carrousel := 70;
                           END_IF;

                           //Popup 1 TO PopUp 2 conveyors
                           IF #Source_Location_Carousel.Device_Type = 15 AND #Destination_Location_Carousel.Device_Type = 16 AND
                               "Control_DB".PopUp_Cnv[2].Done AND "Control_DB".PopUp_Cnv[1].Done
                           THEN
                               "Control_DB"."Carrousel_Order Table".SM_State := "Control_DB".PopUp_Cnv[2].SM_State;
                               "Control_DB"."Carrousel_Order Table".Movement_Request_Complete := TRUE;
                               #State_Carrousel := 70;
                           END_IF;

                           //Popup 3 TO PopUp 4 conveyors
                           IF #Source_Location_Carousel.Device_Type = 17 AND #Destination_Location_Carousel.Device_Type = 18 AND
                               "Control_DB".PopUp_Cnv[4].Done AND "Control_DB".PopUp_Cnv[3].Done
                           THEN
                               "Control_DB"."Carrousel_Order Table".SM_State := "Control_DB".PopUp_Cnv[4].SM_State;
                               "Control_DB"."Carrousel_Order Table".Movement_Request_Complete := TRUE;
                               #State_Carrousel := 70;
                           END_IF;

                           //Popup 4 TO Outbound conveyors
                           IF #Source_Location_Carousel.Device_Type = 18 AND #Destination_Location_Carousel.Device_Type = 14 AND
                               "Control_DB".Outbound_Cnv.Done AND "Control_DB".PopUp_Cnv[4].Done
                           THEN
                               "Control_DB"."Carrousel_Order Table".SM_State := "Control_DB".Outbound_Cnv.SM_State;
                               "Control_DB"."Carrousel_Order Table".Movement_Request_Complete := TRUE;
                               #State_Carrousel := 70;
                           END_IF;

                       70: //Wait for the ACK before we go back to Idle
                               //Inbound to popup 1 conveyors
                           IF #Source_Location_Carousel.Device_Type = 13 AND #Destination_Location_Carousel.Device_Type = 15
                           THEN
                               "Control_DB"."Carrousel_Order Table".SM_State := "Control_DB".PopUp_Cnv[1].SM_State;

                               //Popup 1 TO PopUp 2 conveyors
                           ELSIF #Source_Location_Carousel.Device_Type = 15 AND #Destination_Location_Carousel.Device_Type = 16
                           THEN
                               "Control_DB"."Carrousel_Order Table".SM_State := "Control_DB".PopUp_Cnv[2].SM_State;

                               //Popup 3 TO PopUp 4 conveyors
                           ELSIF #Source_Location_Carousel.Device_Type = 17 AND #Destination_Location_Carousel.Device_Type = 18
                           THEN
                               "Control_DB"."Carrousel_Order Table".SM_State := "Control_DB".PopUp_Cnv[4].SM_State;

                               //Popup 4 TO Outbound conveyors
                           ELSIF #Source_Location_Carousel.Device_Type = 18 AND #Destination_Location_Carousel.Device_Type = 14
                           THEN
                               "Control_DB"."Carrousel_Order Table".SM_State := "Control_DB".Outbound_Cnv.SM_State;
                           END_IF;

                           IF "Control_DB"."Carrousel_Order Table".Movement_Request_Complete_Ack THEN
                               #State_Carrousel := 250;
                           END_IF;

                           //=========================== Transfer Pallet Chain to Chain  ===========================

